	n_PHASE_LOWER:
		lr_ToolRz[n_Robot] := lr_ToolRz[n_Robot] * (1.0 - MIN(1.0, lr_Dt * 5.0));
		IF n_Robot = 1 THEN
			lr_TiltRx := _FC_DemoApproach(lr_TiltRx, 0, lr_TILT_SPEED * lr_Dt);
		END_IF
		(* Delta 2 puts the product down straight (both operands are evaluated). *)
		IF m_MoveToward(vio_Tcp := Tcp[n_Robot], vi_lr_TargetX := Tcp[n_Robot].fX, vi_lr_TargetY := Tcp[n_Robot].fY,
			vi_lr_TargetZ := DEMO_GlobalConst.DEMO_lr_BELT_Z + lr_HeldHeight + lr_GripHeight,
			vi_lr_MaxStep := lr_Step)
		AND (n_Robot <> 1 OR lr_TiltRx = 0)
		THEN
			n_Phase[n_Robot] := n_PHASE_RELEASE;
		END_IF

	n_PHASE_RELEASE:
		(* Every carried product is put down where its finger (Delta 3: the flange) holds it. *)
		FOR n_Slot := 0 TO n_HeldCount[n_Robot] - 1 DO
			IF n_HeldBelt[n_Robot, n_Slot] = 0 THEN
				fb_RefBelt REF= fb_Infeed1;
			ELSE
				fb_RefBelt REF= fb_Infeed2;
			END_IF
			(* Put down on the outfeed: it no longer lies on the infeed. *)
			fb_RefBelt.m_RemoveProduct(udn_Held[n_Robot, n_Slot]);
			n_Finger := SEL(n_Robot = 2, n_Slot + 1, 0);
			Grip := m_GripOffset(vi_n_Robot := n_Robot, vi_n_Finger := n_Finger);
			LatchPose.fX := Tcp[n_Robot].fX + Grip.fX;
			LatchPose.fY := Tcp[n_Robot].fY + Grip.fY;
			LatchPose.fZ := DEMO_GlobalConst.DEMO_lr_BELT_Z;
			(* A product carried at a finger keeps the finger's turn; one at the flange is turned with the base. *)
			LatchPose.fRz := SEL(n_Robot = 2, lr_ToolRz[n_Robot], 0);
			IF fb_Outfeed.m_LatchProduct(vi_udn_Id := DEMO_GlobalVar.DEMO_udn_NextId,
				vi_LatchPose := fb_Outfeed.m_McsToBelt(vi_Pose := LatchPose),
				vi_udn_ProductType := udn_HeldType[n_Robot, n_Slot], vi_lr_LatchBeltPosition := 0,
				vi_b_UseLatchBeltPosition := FALSE, vi_e_State := E_VisuProductState.PLACED,
				vi_udn_ClientId := fb_RefRobot.m_Id())
			THEN
				(* A sample stays marked on the outfeed. *)
				fb_Outfeed.m_SetProductMark(vi_udn_Id := DEMO_GlobalVar.DEMO_udn_NextId, vi_un_Mark := un_HeldMark[n_Robot, n_Slot]);
				DEMO_GlobalVar.DEMO_udn_NextId := DEMO_GlobalVar.DEMO_udn_NextId + 1;
			END_IF
			udn_Held[n_Robot, n_Slot] := 0;
		END_FOR
		n_HeldCount[n_Robot] := 0;
		un_Placed[n_Robot] := un_Placed[n_Robot] + 1;
		n_Phase[n_Robot] := n_PHASE_IDLE;
END_CASE
m_Sequence := TRUE;
END_METHOD

(****************************************************************************************************<br>
© Syntegon Group.<br>
All rights reserved, also regarding any disposal, exploitation, reproduction, editing, distribution,<br>
as well as in the event of applications for industrial property rights.<br>
*****************************************************************************************************<br>
DESCRIPTION:<br>
Follows the current target of Delta n_Robot by its id (register indices shift when entries are removed),<br>
selects its infeed into fb_RefBelt and the finger used for the current pick into n_Finger and Grip. Sets the height<br>
of the product carried or approached and the Delta 3 finger distance closed around it.<br>
****************************************************************************************************)
METHOD PRIVATE m_Target : BOOL
VAR
	lr_TempHalfLength					: LREAL;	// [mm]
	lr_TempHalfWidth					: LREAL;	// [mm]
	lr_TempRadius						: LREAL;	// [mm] corner radius of a rounded box
	lr_TempOuter						: LREAL;	// [mm] radius of the circle around the product's outline
END_VAR
(* Current target *)
b_Found := FALSE;
IF udn_TargetId[n_Robot] <> 0 THEN
	IF n_TargetBelt[n_Robot] = 0 THEN
		fb_RefBelt REF= fb_Infeed1;
	ELSE
		fb_RefBelt REF= fb_Infeed2;
	END_IF
	IF fb_RefBelt.m_FindProduct(udn_TargetId[n_Robot]) >= 0 THEN
		b_Found := fb_RefBelt.m_GetProduct(vi_un_Index := INT_TO_UINT(fb_RefBelt.m_FindProduct(udn_TargetId[n_Robot])),
			vo_Product => Product, vo_Pose => ProductPose);
	END_IF
END_IF

(* Only approaching and descending follow a target; carried products are tracked in udn_Held. *)
IF (n_Phase[n_Robot] = n_PHASE_APPROACH OR n_Phase[n_Robot] = n_PHASE_DESCEND) AND NOT b_Found THEN
	n_Phase[n_Robot] := n_PHASE_IDLE;
	udn_TargetId[n_Robot] := 0;
END_IF
IF b_Found THEN
	ProductPose := fb_RefBelt.m_BeltToMcs(vi_Pose := ProductPose);
	lr_X := ProductPose.fX + lr_LEAD;
	lr_Y := ProductPose.fY;
	lr_TopZ := ProductPose.fZ + lr_TYPE_HEIGHT[LIMIT(1, Product.nProductType, udn_TYPE_COUNT)];
	lr_TargetRz := ProductPose.fRz;
END_IF

(* Size of the product carried, else of the one approached: Delta 1 carries a pair of one type, so its first slot
   stands for both. *)
IF n_HeldCount[n_Robot] > 0 THEN
	udn_Type := LIMIT(1, udn_HeldType[n_Robot, 0], udn_TYPE_COUNT);
ELSIF b_Found THEN
	udn_Type := LIMIT(1, Product.nProductType, udn_TYPE_COUNT);
ELSE
	udn_Type := 1;
END_IF
lr_HeldHeight := lr_TYPE_HEIGHT[udn_Type];
(* Delta 3 closes its fingers on a circle just around the product's outline: around a box's corners, a cylinder's
   larger radius, or a rounded box's corner arcs. *)
lr_TempHalfLength := lr_TYPE_LENGTH[udn_Type] / 2.0;
lr_TempHalfWidth := lr_TYPE_WIDTH[udn_Type] / 2.0;
CASE e_TYPE_SHAPE[udn_Type] OF
	E_VisuProductShape.CYLINDER:
		lr_TempOuter := MAX(lr_TempHalfLength, lr_TempHalfWidth);
	E_VisuProductShape.ROUNDED_BOX:
		lr_TempRadius := MIN(lr_TYPE_CORNER_RADIUS[udn_Type], MIN(lr_TempHalfLength, lr_TempHalfWidth));
		lr_TempOuter := SQRT((lr_TempHalfLength - lr_TempRadius) * (lr_TempHalfLength - lr_TempRadius)
							+ (lr_TempHalfWidth - lr_TempRadius) * (lr_TempHalfWidth - lr_TempRadius)) + lr_TempRadius;
ELSE
	lr_TempOuter := SQRT(lr_TempHalfLength * lr_TempHalfLength + lr_TempHalfWidth * lr_TempHalfWidth);
END_CASE
lr_SpreadClosed := lr_TempOuter + lr_RING_CLEARANCE;

(* Finger used for the current pick: Delta 1 fills its cups one after the other, Delta 3 carries at the flange
   between its fingers. *)
CASE n_Robot OF
	0:
		n_Finger := MIN(n_HeldCount[n_Robot] + 1, 2);
		lr_GripHeight := DEMO_GlobalConst.DEMO_lr_CUP_HEIGHT;
	1:
		n_Finger := 1;
		lr_GripHeight := lr_TILT_HEIGHT;
ELSE
	n_Finger := 0;
	lr_GripHeight := 0;
END_CASE
Grip := m_GripOffset(vi_n_Robot := n_Robot, vi_n_Finger := n_Finger);
m_Target := b_Found;
END_METHOD

(****************************************************************************************************<br>
© Syntegon Group.<br>
All rights reserved, also regarding any disposal, exploitation, reproduction, editing, distribution,<br>
as well as in the event of applications for industrial property rights.<br>
*****************************************************************************************************<br>
DESCRIPTION:<br>
The demo's tracking of Vision 1: latches a raw detection on Infeed 1 at the belt position it was seen at, as<br>
Vision 1's, and marks every tenth product as a sample.<br>
*****************************************************************************************************<br>
OUTPUT VALUES:<br>
TRUE if the product entered the register.<br>
****************************************************************************************************)
METHOD PRIVATE m_Track : BOOL
VAR_INPUT
	vi_Detection						: TVisuDemo_Detection;	// from the product generator
END_VAR
m_Track := fb_Infeed1.m_LatchProduct(vi_udn_Id := DEMO_GlobalVar.DEMO_udn_NextId,
	vi_LatchPose := fb_Infeed1.m_McsToBelt(vi_Pose := vi_Detection.Pose),
	vi_udn_ProductType := vi_Detection.udn_ProductType, vi_lr_LatchBeltPosition := vi_Detection.lr_BeltPosition,
	vi_b_UseLatchBeltPosition := TRUE, vi_e_State := E_VisuProductState.DETECTED, vi_udn_ClientId := fb_Vision1.m_Id());
IF m_Track THEN
	un_Vision1Latches := un_Vision1Latches + 1;
	IF un_Vision1Latches MOD un_SAMPLE_EVERY = 0 THEN
		fb_Infeed1.m_SetProductMark(vi_udn_Id := DEMO_GlobalVar.DEMO_udn_NextId, vi_un_Mark := un_SAMPLE_MARK);
	END_IF
	DEMO_GlobalVar.DEMO_udn_NextId := DEMO_GlobalVar.DEMO_udn_NextId + 1;
END_IF
END_METHOD

END_PROGRAM

// ---- POUs/P_VisuDemoFxx.TcPOU
(****************************************************************************************************<br>
© Syntegon Group.<br>
All rights reserved, also regarding any disposal, exploitation, reproduction, editing, distribution,<br>
as well as in the event of applications for industrial property rights.<br>
*****************************************************************************************************<br>
DESCRIPTION:<br>
DEMO ONLY: Fxx application (Y = 2500). Products arrive irregularly on the Fxx infeed; an XTS loop above the belts<br>
takes them over and puts them onto the Fxx outfeed with an even spacing. Mover 3 and the first far curve module<br>
are in a fault now and then. The Fxx outfeed is a conveyor without a body.<br>
Called by P_VisuDemo.<br>
****************************************************************************************************)
PROGRAM P_VisuDemoFxx
VAR
	fb_FxxInfeed						: _FB_VisuConveyor;
	fb_FxxOutfeed						: _FB_VisuConveyor;
	fb_Fxx								: _FB_VisuXtsLoop;

	(* Conveyors *)
	lr_Dt								: LREAL;	// [s] cycle time
	udn_Seed							: UDINT := 23456;	// [-] pseudo random generator state
	lr_InfeedPosition					: LREAL;	// [mm] belt position of the Fxx infeed
	lr_OutfeedPosition					: LREAL;	// [mm] belt position of the Fxx outfeed
	lr_SinceSpawn						: LREAL;	// [s] since the last product
	lr_SpawnInterval					: LREAL := 0.6;	// [s] irregular: the Fxx evens the gaps out
	BeltPose							: ST_VisuPose;
	LatchPose							: ST_VisuPlanarPose;
	XtsPose								: ST_VisuPose;

	(* XTS loop: unwrapped track position per mover; queued movers wait just before the perimeter (= 0). *)
	b_LoopInitialised					: BOOL;
	lr_LoopS							: ARRAY[0..11] OF LREAL;	// [mm] per mover (n_LOOP_MOVERS)
	n_LoopMode							: ARRAY[0..11] OF INT;
	udn_LoopProduct						: ARRAY[0..11] OF UDINT;	// [-] product id on the Fxx infeed
	MoverFingers						: ARRAY[0..VISU_GlobalConst_Param.VISU_un_MAX_FINGERS - 1] OF ST_VisuFingerState;	// the mover's cup: grips
	un_Module							: UINT;	// [-] track module being set
	e_ModuleKind						: E_VisuModuleKind;
END_VAR
VAR CONSTANT
	lr_FXX_Y							: LREAL := 2500;	// [mm]
	lr_FXX_INFEED_LENGTH				: LREAL := 2000;	// [mm]
	lr_FXX_INFEED_SPEED					: LREAL := 150;	// [mm/s]
	lr_FXX_OUTFEED_X					: LREAL := 2400;	// [mm]
	lr_FXX_OUTFEED_LENGTH				: LREAL := 3000;	// [mm]
	lr_FXX_OUTFEED_SPEED				: LREAL := 300;	// [mm/s]
	lr_LOOP_X							: LREAL := 1000;	// [mm] start of the lower straight above the Fxx infeed
	un_LOOP_STRAIGHT_MODULES			: UINT := 10;	// [-] straight XTS modules per side, joined at each end by two left curve modules
	lr_LOOP_TOOL_OFFSET					: LREAL := 120;	// [mm]
	n_LOOP_MOVERS						: INT := 12;	// [-] size of the lr_LoopS, n_LoopMode and udn_LoopProduct arrays
	lr_LOOP_SLOT						: LREAL := 130;	// [mm] queue spacing
	lr_LOOP_GRIP						: LREAL := 300;	// [mm] track position where the product is gripped
	lr_LOOP_RELEASE						: LREAL := 600;	// [mm] track position where the mover stops following the infeed
	lr_LOOP_PLACE						: LREAL := 2000;	// [mm] track position of the hand-over to the Fxx outfeed
	lr_LOOP_DELIVER_SPEED				: LREAL := 700;	// [mm/s]
	lr_LOOP_RETURN_SPEED				: LREAL := 900;	// [mm/s]
	lr_FAULT_START						: LREAL := 10;	// [s] start of the mover 3 fault in the fault period
	lr_MODULE_FAULT_START				: LREAL := 15;	// [s] start of the fault of the first far curve module
	n_LOOP_QUEUE						: INT := 0;
	n_LOOP_TRACK						: INT := 1;
	n_LOOP_DELIVER						: INT := 2;
	n_LOOP_RETURN						: INT := 3;
END_VAR

lr_Dt := DEMO_GlobalVar.DEMO_lr_Dt;


(****************************************************************************************************)
(* REGISTRATION (idempotent, every cycle)                                                           *)
(****************************************************************************************************)
fb_FxxInfeed.m_Register(vio_Manifest := GVL_Visu.stManifest, vi_udn_Id := 4, vi_str_Name := 'Fxx infeed');
fb_FxxOutfeed.m_Register(vio_Manifest := GVL_Visu.stManifest, vi_udn_Id := 5, vi_str_Name := 'Fxx outfeed');
fb_Fxx.m_Register(vio_Manifest := GVL_Visu.stManifest, vi_udn_Id := 20, vi_str_Name := 'Fxx');


(****************************************************************************************************)
(* CONVEYORS (configuration idempotent, every cycle)                                                *)
(****************************************************************************************************)
BeltPose.fX := 0;
BeltPose.fY := lr_FXX_Y;
BeltPose.fZ := DEMO_GlobalConst.DEMO_lr_BELT_Z;
fb_FxxInfeed.m_SetPose(vi_Pose := BeltPose);
fb_FxxInfeed.m_Configure(vi_lr_Length := lr_FXX_INFEED_LENGTH,
	vi_lr_Width := DEMO_GlobalConst.DEMO_lr_BELT_WIDTH);
BeltPose.fX := lr_FXX_OUTFEED_X;
(* The outfeed's coordinate system lies on its right edge (seen in the conveying direction). *)
fb_FxxOutfeed.m_SetOriginShift(vi_lr_X := 0, vi_lr_Y := -DEMO_GlobalConst.DEMO_lr_BELT_WIDTH / 2, vi_lr_Z := 0);
fb_FxxOutfeed.m_SetPose(vi_Pose := BeltPose);
fb_FxxOutfeed.m_Configure(vi_lr_Length := lr_FXX_OUTFEED_LENGTH,
	vi_lr_Width := DEMO_GlobalConst.DEMO_lr_BELT_WIDTH);
(* A conveyor without a body: only its products, zones and axis (from the shifted origin) are drawn. *)
fb_FxxOutfeed.m_SetBodyVisible(vi_b_Visible := FALSE);
fb_FxxInfeed.m_SetProductType(vi_udn_Id := 1, vi_lr_Length := DEMO_GlobalConst.DEMO_lr_PRODUCT_LENGTH,
	vi_lr_Width := DEMO_GlobalConst.DEMO_lr_PRODUCT_WIDTH, vi_lr_Height := DEMO_GlobalConst.DEMO_lr_PRODUCT_HEIGHT,
	vi_e_Shape := E_VisuProductShape.BOX, vi_lr_CornerRadius := 0);
fb_FxxOutfeed.m_SetProductType(vi_udn_Id := 1, vi_lr_Length := DEMO_GlobalConst.DEMO_lr_PRODUCT_LENGTH,
	vi_lr_Width := DEMO_GlobalConst.DEMO_lr_PRODUCT_WIDTH, vi_lr_Height := DEMO_GlobalConst.DEMO_lr_PRODUCT_HEIGHT,
	vi_e_Shape := E_VisuProductShape.BOX, vi_lr_CornerRadius := 0);

(* Belt travel *)
lr_InfeedPosition := lr_InfeedPosition + lr_FXX_INFEED_SPEED * lr_Dt;
lr_OutfeedPosition := lr_OutfeedPosition + lr_FXX_OUTFEED_SPEED * lr_Dt;
fb_FxxInfeed.m_SetBeltPosition(lr_InfeedPosition);
fb_FxxOutfeed.m_SetBeltPosition(lr_OutfeedPosition);


(****************************************************************************************************)
(* PRODUCT INFEED: irregular gaps                                                                   *)
(****************************************************************************************************)
lr_SinceSpawn := lr_SinceSpawn + lr_Dt;
IF lr_SinceSpawn >= lr_SpawnInterval THEN
	lr_SinceSpawn := 0;
	udn_Seed := udn_Seed * 1103515245 + 12345;
	lr_SpawnInterval := 0.4 + UDINT_TO_LREAL(udn_Seed MOD 1000) / 1000.0 * 1.2;
	LatchPose.fX := 100;
	LatchPose.fY := lr_FXX_Y;
	LatchPose.fZ := DEMO_GlobalConst.DEMO_lr_BELT_Z;
	LatchPose.fRz := 0;
	IF fb_FxxInfeed.m_LatchProduct(vi_udn_Id := DEMO_GlobalVar.DEMO_udn_NextId,
		vi_LatchPose := fb_FxxInfeed.m_McsToBelt(vi_Pose := LatchPose),
		vi_udn_ProductType := 1, vi_lr_LatchBeltPosition := 0, vi_b_UseLatchBeltPosition := FALSE,
		vi_e_State := E_VisuProductState.DETECTED, vi_udn_ClientId := 0)
	THEN
		DEMO_GlobalVar.DEMO_udn_NextId := DEMO_GlobalVar.DEMO_udn_NextId + 1;
	END_IF
END_IF


(****************************************************************************************************)
(* XTS LOOP                                                                                         *)
(****************************************************************************************************)
XtsPose.fX := lr_LOOP_X;
XtsPose.fY := lr_FXX_Y;
XtsPose.fZ := DEMO_GlobalConst.DEMO_lr_BELT_Z + DEMO_GlobalConst.DEMO_lr_PRODUCT_HEIGHT + lr_LOOP_TOOL_OFFSET;
XtsPose.fRz := 0;
(* The flange sits one cup height closer to the track, so the cup's grip point is at the products' tops. *)
fb_Fxx.m_SetPose(vi_Pose := XtsPose);
fb_Fxx.m_Configure(vi_lr_ToolOffset := lr_LOOP_TOOL_OFFSET - DEMO_GlobalConst.DEMO_lr_CUP_HEIGHT,
	vi_lr_MoverLength := 100, vi_lr_MoverWidth := 60);
(* Track: per side the straight modules, then two left curve modules turning up and back. *)
FOR un_Module := 1 TO 2 * (un_LOOP_STRAIGHT_MODULES + 2) DO
	IF (un_Module - 1) MOD (un_LOOP_STRAIGHT_MODULES + 2) < un_LOOP_STRAIGHT_MODULES THEN
		e_ModuleKind := E_VisuModuleKind.STRAIGHT;
	ELSE
		e_ModuleKind := E_VisuModuleKind.CURVE_LEFT;
	END_IF
	fb_Fxx.m_SetModule(vi_un_Module := un_Module, vi_e_Kind := e_ModuleKind,
		vi_lr_Length := VISU_GlobalConst.VISU_lr_XTS_MODULE_LENGTH);
END_FOR
fb_Fxx.m_SetModuleFault(vi_un_Module := un_LOOP_STRAIGHT_MODULES + 1,
	vi_b_Fault := DEMO_GlobalVar.DEMO_lr_FaultPhase >= lr_MODULE_FAULT_START
					AND DEMO_GlobalVar.DEMO_lr_FaultPhase < lr_MODULE_FAULT_START + DEMO_GlobalConst.DEMO_lr_FAULT_DURATION,
	vi_str_FaultMessage := 'Overtemperature');
fb_Fxx.m_SetFinger(vi_un_Finger := 1, vi_lr_Diameter := DEMO_GlobalConst.DEMO_lr_CUP_DIAMETER,
	vi_lr_Height := DEMO_GlobalConst.DEMO_lr_CUP_HEIGHT);
(* The cup hangs at the flange centre; the movers report no finger poses, the visualisation places the cup by its
   offset on every mover's flange (ADR 0018). *)
fb_Fxx.m_SetFingerOffset(vi_un_Finger := 1, vi_lr_X := 0, vi_lr_Y := 0, vi_lr_Z := 0, vi_lr_Rz := 0);
fb_Fxx.m_SetFingersOnFlange(vi_b_OnFlange := TRUE);
fb_Fxx.m_SetZone(vi_un_Zone := 1, vi_udn_ConveyorId := fb_FxxInfeed.m_Id(), vi_lr_Start := lr_LOOP_X,
	vi_lr_End := lr_LOOP_X + lr_LOOP_RELEASE, vi_lr_AllocationOffset := 0, vi_lr_CcsOffset := lr_LOOP_X,
	vi_lr_StartY := 0, vi_lr_EndY := 0);
fb_Fxx.m_SetZone(vi_un_Zone := 2, vi_udn_ConveyorId := fb_FxxOutfeed.m_Id(),
	vi_lr_Start := lr_LOOP_X + lr_LOOP_PLACE - lr_FXX_OUTFEED_X - 300,
	vi_lr_End := lr_LOOP_X + lr_LOOP_PLACE - lr_FXX_OUTFEED_X + 100,
	vi_lr_AllocationOffset := 0, vi_lr_CcsOffset := lr_LOOP_X + lr_LOOP_PLACE - lr_FXX_OUTFEED_X,
	vi_lr_StartY := 0, vi_lr_EndY := 0);
m_Step();


(****************************************************************************************************)
(* HOUSEKEEPING                                                                                     *)
(****************************************************************************************************)
fb_FxxInfeed.m_RemoveProductsBeyond(lr_FXX_INFEED_LENGTH + DEMO_GlobalConst.DEMO_lr_REMOVE_BEYOND_END);
fb_FxxOutfeed.m_RemoveProductsBeyond(lr_FXX_OUTFEED_LENGTH + DEMO_GlobalConst.DEMO_lr_REMOVE_BEYOND_END);

(****************************************************************************************************<br>
© Syntegon Group.<br>
All rights reserved, also regarding any disposal, exploitation, reproduction, editing, distribution,<br>
as well as in the event of applications for industrial property rights.<br>
*****************************************************************************************************<br>
DESCRIPTION:<br>
XTS loop: the queue head takes over the next product arriving on the Fxx infeed under the start of the lower<br>
straight, follows it, grips it, carries it faster to the Fxx outfeed and releases it there; the mover then<br>
runs round to the queue.<br>
****************************************************************************************************)
METHOD PRIVATE m_Step : BOOL
VAR
	lr_TempPerimeter					: LREAL;	// [mm]
	lr_TempS							: LREAL;	// [mm]
	lr_TempX							: LREAL;	// [mm]
	lr_TempRz							: LREAL;	// [deg]
	n_TempI								: INT;
	n_TempJ								: INT;
	n_TempRank							: INT;
	n_TempHead							: INT;
	b_TempHeadReady						: BOOL;
	lr_TempMinTrack						: LREAL;	// [mm]
	n_TempIdx							: INT;
	un_TempIndex						: UINT;
	TempProduct							: ST_VisuProduct;
	TempPose							: ST_VisuPlanarPose;
	TempLatch							: ST_VisuPlanarPose;
END_VAR
(****************************************************************************************************)
(* QUEUE AND TAKE-OVER                                                                              *)
(****************************************************************************************************)
lr_TempPerimeter := fb_Fxx.m_TrackLength();
IF NOT b_LoopInitialised THEN
	FOR n_TempI := 0 TO n_LOOP_MOVERS - 1 DO
		lr_LoopS[n_TempI] := lr_TempPerimeter - INT_TO_LREAL(n_TempI) * lr_LOOP_SLOT;
		n_LoopMode[n_TempI] := n_LOOP_QUEUE;
	END_FOR
	b_LoopInitialised := TRUE;
END_IF

(* Queued movers close up towards their slots before the start of the lower straight. *)
n_TempHead := -1;
FOR n_TempI := 0 TO n_LOOP_MOVERS - 1 DO
	IF n_LoopMode[n_TempI] = n_LOOP_QUEUE THEN
		n_TempRank := 0;
		FOR n_TempJ := 0 TO n_LOOP_MOVERS - 1 DO
			IF n_LoopMode[n_TempJ] = n_LOOP_QUEUE
			AND (lr_LoopS[n_TempJ] > lr_LoopS[n_TempI] OR (lr_LoopS[n_TempJ] = lr_LoopS[n_TempI] AND n_TempJ < n_TempI))
			THEN
				n_TempRank := n_TempRank + 1;
			END_IF
		END_FOR
		lr_LoopS[n_TempI] := MIN(lr_LoopS[n_TempI] + lr_LOOP_RETURN_SPEED * lr_Dt,
								lr_TempPerimeter - INT_TO_LREAL(n_TempRank) * lr_LOOP_SLOT);
		IF n_TempRank = 0 THEN
			n_TempHead := n_TempI;
		END_IF
	END_IF
END_FOR

(* The queue head takes over the next product arriving under the start of the lower straight.
   ST evaluates both operands of AND, so the index check must be a separate IF (head = -1: queue empty). *)
b_TempHeadReady := FALSE;
IF n_TempHead >= 0 THEN
	b_TempHeadReady := lr_LoopS[n_TempHead] >= lr_TempPerimeter - 1;
END_IF
(* Movers cannot overlap: the next product must be at least one slot behind the last mover following one. *)
lr_TempMinTrack := 1.0E9;
FOR n_TempI := 0 TO n_LOOP_MOVERS - 1 DO
	IF n_LoopMode[n_TempI] = n_LOOP_TRACK THEN
		lr_TempMinTrack := MIN(lr_TempMinTrack, lr_LoopS[n_TempI]);
	END_IF
END_FOR
IF b_TempHeadReady THEN
	un_TempIndex := 0;
	WHILE n_LoopMode[n_TempHead] = n_LOOP_QUEUE AND un_TempIndex < fb_FxxInfeed.m_ProductCount() DO
		fb_FxxInfeed.m_GetProduct(vi_un_Index := un_TempIndex, vo_Product => TempProduct, vo_Pose => TempPose);
		TempPose := fb_FxxInfeed.m_BeltToMcs(vi_Pose := TempPose);
		lr_TempX := TempPose.fX - lr_LOOP_X;
		IF TempProduct.eState = E_VisuProductState.DETECTED AND lr_TempX >= 0 AND lr_TempX < lr_LOOP_GRIP
		AND lr_TempMinTrack - lr_TempX >= lr_LOOP_SLOT
		THEN
			fb_FxxInfeed.m_SetProductState(vi_udn_Id := TempProduct.nId, vi_e_State := E_VisuProductState.ASSIGNED,
				vi_udn_ClientId := fb_Fxx.m_Id(), vi_udn_MoverId := INT_TO_UDINT(n_TempHead + 1), vi_udn_FingerId := 0);
			udn_LoopProduct[n_TempHead] := TempProduct.nId;
			n_LoopMode[n_TempHead] := n_LOOP_TRACK;
		END_IF
		un_TempIndex := un_TempIndex + 1;
	END_WHILE
END_IF


(****************************************************************************************************)
(* MOVERS                                                                                           *)
(****************************************************************************************************)
fb_Fxx.m_SetMoverCount(INT_TO_UINT(n_LOOP_MOVERS));
FOR n_TempI := 0 TO n_LOOP_MOVERS - 1 DO
	CASE n_LoopMode[n_TempI] OF
		n_LOOP_TRACK:
			n_TempIdx := fb_FxxInfeed.m_FindProduct(udn_LoopProduct[n_TempI]);
			IF n_TempIdx < 0 THEN
				udn_LoopProduct[n_TempI] := 0;
				n_LoopMode[n_TempI] := n_LOOP_RETURN;
			ELSE
				fb_FxxInfeed.m_GetProduct(vi_un_Index := INT_TO_UINT(n_TempIdx), vo_Product => TempProduct, vo_Pose => TempPose);
				TempPose := fb_FxxInfeed.m_BeltToMcs(vi_Pose := TempPose);
				lr_LoopS[n_TempI] := TempPose.fX - lr_LOOP_X;
				IF lr_LoopS[n_TempI] >= lr_LOOP_GRIP AND TempProduct.eState = E_VisuProductState.ASSIGNED THEN
					fb_FxxInfeed.m_SetProductState(vi_udn_Id := TempProduct.nId, vi_e_State := E_VisuProductState.PICKED,
						vi_udn_ClientId := fb_Fxx.m_Id(), vi_udn_MoverId := INT_TO_UDINT(n_TempI + 1), vi_udn_FingerId := 1);
				END_IF
				IF lr_LoopS[n_TempI] >= lr_LOOP_RELEASE THEN
					n_LoopMode[n_TempI] := n_LOOP_DELIVER;
				END_IF
			END_IF

		n_LOOP_DELIVER:
			lr_LoopS[n_TempI] := MIN(lr_LoopS[n_TempI] + lr_LOOP_DELIVER_SPEED * lr_Dt, lr_LOOP_PLACE);
			IF lr_LoopS[n_TempI] >= lr_LOOP_PLACE THEN
				lr_TempRz := 0;
				n_TempIdx := fb_FxxInfeed.m_FindProduct(udn_LoopProduct[n_TempI]);
				IF n_TempIdx >= 0 THEN
					fb_FxxInfeed.m_GetProduct(vi_un_Index := INT_TO_UINT(n_TempIdx), vo_Product => TempProduct, vo_Pose => TempPose);
					lr_TempRz := TempProduct.stLatchPose.fRz;
					(* Put down on the outfeed: it no longer lies on the infeed. *)
					fb_FxxInfeed.m_RemoveProduct(TempProduct.nId);
				END_IF
				TempLatch.fX := lr_LOOP_X + lr_LoopS[n_TempI];
				TempLatch.fY := lr_FXX_Y;
				TempLatch.fZ := DEMO_GlobalConst.DEMO_lr_BELT_Z;
				TempLatch.fRz := lr_TempRz;
				IF fb_FxxOutfeed.m_LatchProduct(vi_udn_Id := DEMO_GlobalVar.DEMO_udn_NextId,
					vi_LatchPose := fb_FxxOutfeed.m_McsToBelt(vi_Pose := TempLatch),
					vi_udn_ProductType := 1, vi_lr_LatchBeltPosition := 0, vi_b_UseLatchBeltPosition := FALSE,
					vi_e_State := E_VisuProductState.PLACED, vi_udn_ClientId := fb_Fxx.m_Id())
				THEN
					DEMO_GlobalVar.DEMO_udn_NextId := DEMO_GlobalVar.DEMO_udn_NextId + 1;
				END_IF
				udn_LoopProduct[n_TempI] := 0;
				n_LoopMode[n_TempI] := n_LOOP_RETURN;
			END_IF

		n_LOOP_RETURN:
			lr_LoopS[n_TempI] := lr_LoopS[n_TempI] + lr_LOOP_RETURN_SPEED * lr_Dt;
			IF lr_LoopS[n_TempI] >= lr_TempPerimeter - INT_TO_LREAL(n_LOOP_MOVERS) * lr_LOOP_SLOT THEN
				n_LoopMode[n_TempI] := n_LOOP_QUEUE;
			END_IF
	END_CASE

	(* Report the mover with its cup: whether it grips; its pose follows from its offset on the flange. *)
	lr_TempS := lr_LoopS[n_TempI];
	IF lr_TempS >= lr_TempPerimeter THEN
		lr_TempS := lr_TempS - lr_TempPerimeter;
	END_IF
	MoverFingers[0].bActive := n_LoopMode[n_TempI] = n_LOOP_DELIVER
							OR (n_LoopMode[n_TempI] = n_LOOP_TRACK AND lr_LoopS[n_TempI] >= lr_LOOP_GRIP);

	(* Demo fault: mover 3 now and then. *)
	fb_Fxx.m_SetMover(vi_un_Index := INT_TO_UINT(n_TempI), vi_udn_Id := INT_TO_UDINT(n_TempI + 1), vi_lr_Position := lr_TempS,
		vi_FingerStates := MoverFingers,
		vi_b_Fault := n_TempI = 2 AND DEMO_GlobalVar.DEMO_lr_FaultPhase >= lr_FAULT_START
					AND DEMO_GlobalVar.DEMO_lr_FaultPhase < lr_FAULT_START + DEMO_GlobalConst.DEMO_lr_FAULT_DURATION,
		vi_str_FaultMessage := 'Following error');
END_FOR
m_Step := TRUE;
END_METHOD

END_PROGRAM

// ---- POUs/P_VisuDemoIdh.TcPOU
(****************************************************************************************************<br>
© Syntegon Group.<br>
All rights reserved, also regarding any disposal, exploitation, reproduction, editing, distribution,<br>
as well as in the event of applications for industrial property rights.<br>
*****************************************************************************************************<br>
DESCRIPTION:<br>
DEMO ONLY: IDH application (Y = 4100..4850). An XTS gantry with four movers picks products from the IDH infeed<br>
in batches and places them onto the tray belt. Mover 2 is in a fault now and then. Called by P_VisuDemo.<br>
****************************************************************************************************)
PROGRAM P_VisuDemoIdh
VAR
	fb_IdhInfeed						: _FB_VisuConveyor;
	fb_IdhTray							: _FB_VisuConveyor;
	fb_Idh								: _FB_VisuXtsGantry;
	(* Syn_Config (ADR 0017): the IDH runs with the parameter set the configurator writes (pose, track, zones,
	   gripper, limit areas), else with its program values; taken over at once in the demo. The simulated motion keeps to the
	   program's track. *)
	fb_IdhParam							: SynConfig._FB_ConfigXtsGantry;
	IdhDefault							: SynConfig.ST_ConfigXtsGantryParam;	// program values of the IDH

	(* Conveyors *)
	lr_Dt								: LREAL;	// [s] cycle time
	udn_Seed							: UDINT := 34567;	// [-] pseudo random generator state
	lr_InfeedPosition					: LREAL;	// [mm] belt position of the IDH infeed
	lr_TrayPosition						: LREAL;	// [mm] belt position of the tray belt
	lr_SinceSpawn						: LREAL;	// [s] since the last product
	lr_SpawnInterval					: LREAL := 0.8;	// [s]
	BeltPose							: ST_VisuPose;
	LatchPose							: ST_VisuPlanarPose;

	(* XTS gantry *)
	n_GantryPhase						: INT;
	lr_GantryZ							: LREAL;	// [mm]
	lr_GantryWait						: ARRAY[0..3] OF LREAL := [100, 300, 500, 700];	// [mm]
	lr_GantryPos						: ARRAY[0..3] OF LREAL := [100, 300, 500, 700];	// [mm]
	lr_GantryX							: ARRAY[0..3] OF LREAL := [200, 200, 200, 200];	// [mm]
	lr_GantryC							: ARRAY[0..3] OF LREAL;	// [deg]
	b_GantryGrip						: ARRAY[0..3] OF BOOL;
	udn_GantryProduct					: ARRAY[0..3] OF UDINT;	// [-] product id on the IDH infeed
	MoverFingers						: ARRAY[0..VISU_GlobalConst_Param.VISU_un_MAX_FINGERS - 1] OF ST_VisuFingerState;	// the mover's cup
	un_Module							: UINT;	// [-] track module being set
END_VAR
VAR PERSISTENT
	IdhSet								: SynConfig.ST_ConfigXtsGantrySet;	// active parameter set of the IDH, kept over a restart
END_VAR
VAR CONSTANT
	(* Gantry turned by -90 deg: track along MCS +X, X axes towards MCS -Y (IDH infeed under X = 200, tray belt
	   under X = 600). *)
	lr_IDH_INFEED_Y						: LREAL := 4500;	// [mm]
	lr_IDH_INFEED_LENGTH				: LREAL := 4000;	// [mm]
	lr_IDH_INFEED_SPEED					: LREAL := 200;	// [mm/s]
	lr_TRAY_X							: LREAL := 1300;	// [mm]
	lr_TRAY_Y							: LREAL := 4100;	// [mm]
	lr_TRAY_LENGTH						: LREAL := 2000;	// [mm]
	lr_TRAY_SPEED						: LREAL := 80;	// [mm/s]
	lr_GANTRY_X							: LREAL := 1500;	// [mm]
	lr_GANTRY_Y							: LREAL := 4850;	// [mm]
	lr_GANTRY_Z							: LREAL := 1340;	// [mm]
	un_GANTRY_MODULES					: UINT := 6;	// [-]
	lr_GANTRY_MODULE_LENGTH				: LREAL := 250;	// [mm]
	lr_GANTRY_TOOL_X					: LREAL := 150;	// [mm]
	lr_GANTRY_TOOL_Z					: LREAL := -400;	// [mm]
	lr_GANTRY_MOVER_LENGTH				: LREAL := 155;	// [mm]
	lr_GANTRY_GAP						: LREAL := 180;	// [mm] minimum distance between movers
	lr_GANTRY_X_BELT					: LREAL := 200;	// [mm]
	lr_GANTRY_X_TRAY					: LREAL := 600;	// [mm]
	lr_GANTRY_Z_DOWN					: LREAL := -100;	// [mm]
	lr_GANTRY_Z_SPEED					: LREAL := 500;	// [mm/s]
	lr_GANTRY_X_SPEED					: LREAL := 1000;	// [mm/s]
	lr_GANTRY_TRACK_SPEED				: LREAL := 1500;	// [mm/s]
	lr_FAULT_START						: LREAL := 12;	// [s] start of the mover 2 fault in the fault period
	n_GANTRY_COLLECT					: INT := 0;
	n_GANTRY_PICK_DOWN					: INT := 1;
	n_GANTRY_PICK_UP					: INT := 2;
	n_GANTRY_TO_TRAY					: INT := 3;
	n_GANTRY_PLACE_DOWN					: INT := 4;
	n_GANTRY_PLACE_UP					: INT := 5;
	n_GANTRY_RETURN						: INT := 6;
END_VAR

lr_Dt := DEMO_GlobalVar.DEMO_lr_Dt;


(****************************************************************************************************)
(* REGISTRATION (idempotent, every cycle)                                                           *)
(****************************************************************************************************)
fb_IdhInfeed.m_Register(vio_Manifest := GVL_Visu.stManifest, vi_udn_Id := 6, vi_str_Name := 'IDH infeed');
fb_IdhTray.m_Register(vio_Manifest := GVL_Visu.stManifest, vi_udn_Id := 7, vi_str_Name := 'Tray belt');
fb_Idh.m_Register(vio_Manifest := GVL_Visu.stManifest, vi_udn_Id := 30, vi_str_Name := 'IDH');


(****************************************************************************************************)
(* CONVEYORS (configuration idempotent, every cycle)                                                *)
(****************************************************************************************************)
BeltPose.fX := 0;
BeltPose.fY := lr_IDH_INFEED_Y;
BeltPose.fZ := DEMO_GlobalConst.DEMO_lr_BELT_Z;
fb_IdhInfeed.m_SetPose(vi_Pose := BeltPose);
fb_IdhInfeed.m_Configure(vi_lr_Length := lr_IDH_INFEED_LENGTH,
	vi_lr_Width := DEMO_GlobalConst.DEMO_lr_BELT_WIDTH);
BeltPose.fX := lr_TRAY_X;
BeltPose.fY := lr_TRAY_Y;
fb_IdhTray.m_SetPose(vi_Pose := BeltPose);
fb_IdhTray.m_Configure(vi_lr_Length := lr_TRAY_LENGTH, vi_lr_Width := DEMO_GlobalConst.DEMO_lr_BELT_WIDTH);
fb_IdhInfeed.m_SetProductType(vi_udn_Id := 1, vi_lr_Length := DEMO_GlobalConst.DEMO_lr_PRODUCT_LENGTH,
	vi_lr_Width := DEMO_GlobalConst.DEMO_lr_PRODUCT_WIDTH, vi_lr_Height := DEMO_GlobalConst.DEMO_lr_PRODUCT_HEIGHT,
	vi_e_Shape := E_VisuProductShape.BOX, vi_lr_CornerRadius := 0);
fb_IdhTray.m_SetProductType(vi_udn_Id := 1, vi_lr_Length := DEMO_GlobalConst.DEMO_lr_PRODUCT_LENGTH,
	vi_lr_Width := DEMO_GlobalConst.DEMO_lr_PRODUCT_WIDTH, vi_lr_Height := DEMO_GlobalConst.DEMO_lr_PRODUCT_HEIGHT,
	vi_e_Shape := E_VisuProductShape.BOX, vi_lr_CornerRadius := 0);

(* Belt travel *)
lr_InfeedPosition := lr_InfeedPosition + lr_IDH_INFEED_SPEED * lr_Dt;
lr_TrayPosition := lr_TrayPosition + lr_TRAY_SPEED * lr_Dt;
fb_IdhInfeed.m_SetBeltPosition(lr_InfeedPosition);
fb_IdhTray.m_SetBeltPosition(lr_TrayPosition);


(****************************************************************************************************)
(* PRODUCT INFEED: slightly irregular gaps, products turned                                         *)
(****************************************************************************************************)
lr_SinceSpawn := lr_SinceSpawn + lr_Dt;
IF lr_SinceSpawn >= lr_SpawnInterval THEN
	lr_SinceSpawn := 0;
	udn_Seed := udn_Seed * 1103515245 + 12345;
	lr_SpawnInterval := 0.6 + UDINT_TO_LREAL(udn_Seed MOD 1000) / 1000.0 * 0.6;
	LatchPose.fX := 100;
	LatchPose.fY := lr_IDH_INFEED_Y;
	LatchPose.fZ := DEMO_GlobalConst.DEMO_lr_BELT_Z;
	LatchPose.fRz := (UDINT_TO_LREAL((udn_Seed / 1000) MOD 1000) / 1000.0 - 0.5) * 60.0;
	IF fb_IdhInfeed.m_LatchProduct(vi_udn_Id := DEMO_GlobalVar.DEMO_udn_NextId,
		vi_LatchPose := fb_IdhInfeed.m_McsToBelt(vi_Pose := LatchPose),
		vi_udn_ProductType := 1, vi_lr_LatchBeltPosition := 0, vi_b_UseLatchBeltPosition := FALSE,
		vi_e_State := E_VisuProductState.DETECTED, vi_udn_ClientId := 0)
	THEN
		DEMO_GlobalVar.DEMO_udn_NextId := DEMO_GlobalVar.DEMO_udn_NextId + 1;
	END_IF
END_IF


(****************************************************************************************************)
(* XTS GANTRY                                                                                       *)
(****************************************************************************************************)
(* The IDH's program values; its parameter set (Syn_Config) replaces them once the configurator wrote one. Strokes,
   tool offsets and mover size are hardware and stay the program's. *)
IdhDefault.stPose.fX := lr_GANTRY_X;
IdhDefault.stPose.fY := lr_GANTRY_Y;
IdhDefault.stPose.fZ := lr_GANTRY_Z;
IdhDefault.stPose.fRz := -90;
IdhDefault.nModuleCount := un_GANTRY_MODULES;
FOR un_Module := 1 TO un_GANTRY_MODULES DO
	IdhDefault.aModules[un_Module - 1].eKind := E_VisuModuleKind.STRAIGHT;
	IdhDefault.aModules[un_Module - 1].fLength := lr_GANTRY_MODULE_LENGTH;
END_FOR
(* Limit area in the gantry frame (flange coordinates): around the flanges' travel, from over the infeed to over
   the tray belt, along the whole track. *)
IdhDefault.stLimitArea.fXMin := 250;
IdhDefault.stLimitArea.fXMax := 850;
IdhDefault.stLimitArea.fYMin := -50;
IdhDefault.stLimitArea.fYMax := 1550;
IdhDefault.stLimitArea.fZMin := -600;
IdhDefault.stLimitArea.fZMax := -300;
IdhDefault.stLimitArea.bActive := TRUE;
(* Around every mover's flange, cup and product; narrower along the track than the movers' least distance. *)
IdhDefault.stTcpLimitArea.fXMin := -60;
IdhDefault.stTcpLimitArea.fXMax := 60;
IdhDefault.stTcpLimitArea.fYMin := -85;
IdhDefault.stTcpLimitArea.fYMax := 85;
IdhDefault.stTcpLimitArea.fZMin := -100;
IdhDefault.stTcpLimitArea.fZMax := 20;
IdhDefault.stTcpLimitArea.bActive := TRUE;
IdhDefault.nZoneCount := 2;
IdhDefault.aZones[0].nConveyorId := fb_IdhInfeed.m_Id();
IdhDefault.aZones[0].fStart := lr_GANTRY_X;
IdhDefault.aZones[0].fEnd := lr_GANTRY_X + UINT_TO_LREAL(un_GANTRY_MODULES) * lr_GANTRY_MODULE_LENGTH;
IdhDefault.aZones[0].fCcsOffset := lr_GANTRY_X;
IdhDefault.aZones[1].nConveyorId := fb_IdhTray.m_Id();
IdhDefault.aZones[1].fStart := lr_GANTRY_X - lr_TRAY_X;
IdhDefault.aZones[1].fEnd := lr_GANTRY_X - lr_TRAY_X + UINT_TO_LREAL(un_GANTRY_MODULES) * lr_GANTRY_MODULE_LENGTH;
IdhDefault.aZones[1].fCcsOffset := lr_GANTRY_X - lr_TRAY_X;
(* Every mover's suction cup, at the flange centre (ADR 0018); the movers report its live pose, turned by C. It
   comes with the parameter set: the application no longer calls m_SetFinger itself. *)
IdhDefault.nFingerCount := 1;
IdhDefault.aFingers[0].fDiameter := DEMO_GlobalConst.DEMO_lr_CUP_DIAMETER;
IdhDefault.aFingers[0].fHeight := DEMO_GlobalConst.DEMO_lr_CUP_HEIGHT;
fb_IdhParam.m_Register(vio_Manifest := GVL_Config.stManifest, vi_udn_Id := fb_Idh.m_Id());
fb_IdhParam.m_Cycle(vio_Default := IdhDefault, vio_Set := IdhSet, vi_b_ApplyAllowed := TRUE);
fb_Idh.m_Configure(vi_lr_XMin := 0, vi_lr_XMax := 700, vi_lr_ZMin := lr_GANTRY_Z_DOWN, vi_lr_ZMax := 0,
	vi_lr_ToolOffsetX := lr_GANTRY_TOOL_X, vi_lr_ToolOffsetZ := lr_GANTRY_TOOL_Z + DEMO_GlobalConst.DEMO_lr_CUP_HEIGHT,
	vi_lr_MoverLength := lr_GANTRY_MOVER_LENGTH, vi_lr_MoverWidth := 80);
fb_IdhParam.m_PassOn(vio_Visu := fb_Idh);
m_Step();


(****************************************************************************************************)
(* HOUSEKEEPING                                                                                     *)
(****************************************************************************************************)
fb_IdhInfeed.m_RemoveProductsBeyond(lr_IDH_INFEED_LENGTH + DEMO_GlobalConst.DEMO_lr_REMOVE_BEYOND_END);
fb_IdhTray.m_RemoveProductsBeyond(lr_TRAY_LENGTH + DEMO_GlobalConst.DEMO_lr_REMOVE_BEYOND_END);

(****************************************************************************************************<br>
© Syntegon Group.<br>
All rights reserved, also regarding any disposal, exploitation, reproduction, editing, distribution,<br>
as well as in the event of applications for industrial property rights.<br>
*****************************************************************************************************<br>
DESCRIPTION:<br>
Moves the gantry movers along the track: a mover with a product waits at its waiting position until the<br>
product passes underneath and then follows it; a mover without one returns to its waiting position.<br>
Downstream first, so each mover keeps its distance to the one ahead.<br>
****************************************************************************************************)
METHOD PRIVATE m_Follow : BOOL
VAR
	n_TempI								: INT;
	lr_TempGoal							: LREAL;	// [mm]
	lr_TempLimit						: LREAL;	// [mm]
	lr_TempPos							: LREAL;	// [mm]
	lr_TempRz							: LREAL;	// [deg]
END_VAR
FOR n_TempI := 3 TO 0 BY -1 DO
	IF n_TempI = 3 THEN
		lr_TempLimit := UINT_TO_LREAL(un_GANTRY_MODULES) * lr_GANTRY_MODULE_LENGTH - lr_GANTRY_MOVER_LENGTH / 2;
	ELSE
		lr_TempLimit := lr_GantryPos[n_TempI + 1] - lr_GANTRY_GAP;
	END_IF
	lr_TempGoal := lr_GantryWait[n_TempI];
	IF udn_GantryProduct[n_TempI] <> 0 THEN
		IF m_TrackPos(vi_udn_Id := udn_GantryProduct[n_TempI], vo_lr_TrackPos => lr_TempPos, vo_lr_Rz => lr_TempRz) THEN
			lr_TempGoal := MAX(lr_TempPos, lr_GantryWait[n_TempI]);
			(* The cup turns by -90 + C in the MCS (gantry turned by -90 deg), so C = Rz + 90 meets the product. *)
			lr_GantryC[n_TempI] := _FC_DemoApproach(lr_GantryC[n_TempI], lr_TempRz + 90.0, 180.0 * lr_Dt);
		END_IF
	END_IF
	lr_GantryPos[n_TempI] := MIN(_FC_DemoApproach(lr_GantryPos[n_TempI], lr_TempGoal, lr_GANTRY_TRACK_SPEED * lr_Dt),
								lr_TempLimit);
END_FOR
m_Follow := TRUE;
END_METHOD

(****************************************************************************************************<br>
© Syntegon Group.<br>
All rights reserved, also regarding any disposal, exploitation, reproduction, editing, distribution,<br>
as well as in the event of applications for industrial property rights.<br>
*****************************************************************************************************<br>
DESCRIPTION:<br>
XTS gantry: the movers follow up to four products on the IDH infeed (the most downstream mover takes the<br>
first product), then the Z axis lowers all grippers together, the X axes carry the products over the tray<br>
belt, they are put down together and the movers return to their waiting positions.<br>
****************************************************************************************************)
METHOD PRIVATE m_Step : BOOL
VAR
	n_TempI								: INT;
	un_TempIndex						: UINT;
	udn_TempBest						: UDINT;	// [-] product id
	lr_TempBest							: LREAL;	// [mm]
	lr_TempPos							: LREAL;	// [mm]
	lr_TempRz							: LREAL;	// [deg]
	n_TempAssigned						: INT;
	b_TempAllSynced						: BOOL;
	b_TempAnySynced						: BOOL;
	b_TempDone							: BOOL;
	b_TempSynced						: ARRAY[0..3] OF BOOL;
	TempProduct							: ST_VisuProduct;
	TempPose							: ST_VisuPlanarPose;
	TempLatch							: ST_VisuPlanarPose;
END_VAR
(****************************************************************************************************)
(* SEQUENCE                                                                                         *)
(****************************************************************************************************)
CASE n_GantryPhase OF
	n_GANTRY_COLLECT:
		(* Downstream mover first: it takes the most downstream product not yet assigned. *)
		FOR n_TempI := 3 TO 0 BY -1 DO
			IF udn_GantryProduct[n_TempI] = 0 THEN
				udn_TempBest := 0;
				lr_TempBest := -1.0E9;
				FOR un_TempIndex := 1 TO fb_IdhInfeed.m_ProductCount() DO
					fb_IdhInfeed.m_GetProduct(vi_un_Index := un_TempIndex - 1, vo_Product => TempProduct, vo_Pose => TempPose);
					TempPose := fb_IdhInfeed.m_BeltToMcs(vi_Pose := TempPose);
					lr_TempPos := TempPose.fX - lr_GANTRY_X;
					IF TempProduct.eState = E_VisuProductState.DETECTED AND lr_TempPos < lr_GantryPos[n_TempI]
					AND lr_TempPos > -500 AND lr_TempPos > lr_TempBest
					THEN
						udn_TempBest := TempProduct.nId;
						lr_TempBest := lr_TempPos;
					END_IF
				END_FOR
				IF udn_TempBest = 0 THEN
					EXIT;
				END_IF
				fb_IdhInfeed.m_SetProductState(vi_udn_Id := udn_TempBest, vi_e_State := E_VisuProductState.ASSIGNED,
					vi_udn_ClientId := fb_Idh.m_Id(), vi_udn_MoverId := INT_TO_UDINT(n_TempI + 1), vi_udn_FingerId := 0);
				udn_GantryProduct[n_TempI] := udn_TempBest;
			END_IF
		END_FOR
		m_Follow();

		(* Pick once all four are above their products, or at the track end with any of them. *)
		n_TempAssigned := 0;
		b_TempAllSynced := TRUE;
		b_TempAnySynced := FALSE;
		FOR n_TempI := 0 TO 3 DO
			b_TempSynced[n_TempI] := FALSE;
			IF udn_GantryProduct[n_TempI] <> 0 THEN
				n_TempAssigned := n_TempAssigned + 1;
				b_TempSynced[n_TempI] := m_TrackPos(vi_udn_Id := udn_GantryProduct[n_TempI], vo_lr_TrackPos => lr_TempPos,
											vo_lr_Rz => lr_TempRz)
										AND ABS(lr_GantryPos[n_TempI] - lr_TempPos) < 2;
				b_TempAllSynced := b_TempAllSynced AND b_TempSynced[n_TempI];
				b_TempAnySynced := b_TempAnySynced OR b_TempSynced[n_TempI];
			END_IF
		END_FOR
		IF (n_TempAssigned = 4 AND b_TempAllSynced)
		OR (lr_GantryPos[3] >= UINT_TO_LREAL(un_GANTRY_MODULES) * lr_GANTRY_MODULE_LENGTH - 300 AND b_TempAnySynced)
		THEN
			(* Movers not yet above their product give it back. *)
			FOR n_TempI := 0 TO 3 DO
				IF udn_GantryProduct[n_TempI] <> 0 AND NOT b_TempSynced[n_TempI] THEN
					fb_IdhInfeed.m_SetProductState(vi_udn_Id := udn_GantryProduct[n_TempI],
						vi_e_State := E_VisuProductState.DETECTED, vi_udn_ClientId := fb_Idh.m_Id(), vi_udn_MoverId := 0,
						vi_udn_FingerId := 0);
					udn_GantryProduct[n_TempI] := 0;
				END_IF
			END_FOR
			n_GantryPhase := n_GANTRY_PICK_DOWN;
		END_IF

	n_GANTRY_PICK_DOWN:
		m_Follow();
		lr_GantryZ := _FC_DemoApproach(lr_GantryZ, lr_GANTRY_Z_DOWN, lr_GANTRY_Z_SPEED * lr_Dt);
		IF lr_GantryZ = lr_GANTRY_Z_DOWN THEN
			FOR n_TempI := 0 TO 3 DO
				IF udn_GantryProduct[n_TempI] <> 0 THEN
					b_GantryGrip[n_TempI] := TRUE;
					fb_IdhInfeed.m_SetProductState(vi_udn_Id := udn_GantryProduct[n_TempI], vi_e_State := E_VisuProductState.PICKED,
						vi_udn_ClientId := fb_Idh.m_Id(), vi_udn_MoverId := INT_TO_UDINT(n_TempI + 1), vi_udn_FingerId := 1);
				END_IF
			END_FOR
			n_GantryPhase := n_GANTRY_PICK_UP;
		END_IF

	n_GANTRY_PICK_UP:
		lr_GantryZ := _FC_DemoApproach(lr_GantryZ, 0, lr_GANTRY_Z_SPEED * lr_Dt);
		IF lr_GantryZ = 0 THEN
			n_GantryPhase := n_GANTRY_TO_TRAY;
		END_IF

	n_GANTRY_TO_TRAY:
		b_TempDone := TRUE;
		FOR n_TempI := 0 TO 3 DO
			lr_GantryX[n_TempI] := _FC_DemoApproach(lr_GantryX[n_TempI], lr_GANTRY_X_TRAY, lr_GANTRY_X_SPEED * lr_Dt);
			lr_GantryC[n_TempI] := _FC_DemoApproach(lr_GantryC[n_TempI], 0, 180.0 * lr_Dt);
			b_TempDone := b_TempDone AND lr_GantryX[n_TempI] = lr_GANTRY_X_TRAY AND lr_GantryC[n_TempI] = 0;
		END_FOR
		IF b_TempDone THEN
			n_GantryPhase := n_GANTRY_PLACE_DOWN;
		END_IF

	n_GANTRY_PLACE_DOWN:
		lr_GantryZ := _FC_DemoApproach(lr_GantryZ, lr_GANTRY_Z_DOWN, lr_GANTRY_Z_SPEED * lr_Dt);
		IF lr_GantryZ = lr_GANTRY_Z_DOWN THEN
			FOR n_TempI := 0 TO 3 DO
				IF udn_GantryProduct[n_TempI] <> 0 THEN
					(* Put down on the tray: it no longer lies on the infeed. *)
					fb_IdhInfeed.m_RemoveProduct(udn_GantryProduct[n_TempI]);
					(* Turned by -90 deg: gripper at MCS x = track start + position, y = pose y - (X + tool offset). *)
					TempLatch.fX := lr_GANTRY_X + lr_GantryPos[n_TempI];
					TempLatch.fY := lr_GANTRY_Y - (lr_GantryX[n_TempI] + lr_GANTRY_TOOL_X);
					TempLatch.fZ := DEMO_GlobalConst.DEMO_lr_BELT_Z;
					TempLatch.fRz := -90 + lr_GantryC[n_TempI];	// as the cup holds it
					IF fb_IdhTray.m_LatchProduct(vi_udn_Id := DEMO_GlobalVar.DEMO_udn_NextId,
						vi_LatchPose := fb_IdhTray.m_McsToBelt(vi_Pose := TempLatch),
						vi_udn_ProductType := 1, vi_lr_LatchBeltPosition := 0, vi_b_UseLatchBeltPosition := FALSE,
						vi_e_State := E_VisuProductState.PLACED, vi_udn_ClientId := fb_Idh.m_Id())
					THEN
						DEMO_GlobalVar.DEMO_udn_NextId := DEMO_GlobalVar.DEMO_udn_NextId + 1;
					END_IF
					udn_GantryProduct[n_TempI] := 0;
				END_IF
				b_GantryGrip[n_TempI] := FALSE;
			END_FOR
			n_GantryPhase := n_GANTRY_PLACE_UP;
		END_IF

	n_GANTRY_PLACE_UP:
		lr_GantryZ := _FC_DemoApproach(lr_GantryZ, 0, lr_GANTRY_Z_SPEED * lr_Dt);
		IF lr_GantryZ = 0 THEN
			n_GantryPhase := n_GANTRY_RETURN;
		END_IF

	n_GANTRY_RETURN:
		m_Follow();
		b_TempDone := TRUE;
		FOR n_TempI := 0 TO 3 DO
			lr_GantryX[n_TempI] := _FC_DemoApproach(lr_GantryX[n_TempI], lr_GANTRY_X_BELT, lr_GANTRY_X_SPEED * lr_Dt);
			b_TempDone := b_TempDone AND lr_GantryX[n_TempI] = lr_GANTRY_X_BELT AND lr_GantryPos[n_TempI] = lr_GantryWait[n_TempI];
		END_FOR
		IF b_TempDone THEN
			n_GantryPhase := n_GANTRY_COLLECT;
		END_IF
END_CASE


(****************************************************************************************************)
(* REPORT                                                                                           *)
(****************************************************************************************************)
fb_Idh.m_SetZPosition(lr_GantryZ);
fb_Idh.m_SetMoverCount(4);
FOR n_TempI := 0 TO 3 DO
	(* The cup hangs from the flange and turns only about Rz, by the gripper's C. Turned by -90 deg: local (x, y, z)
	   is MCS (gantry x + y, gantry y - x, gantry z + z). *)
	MoverFingers[0].stPose.fX := lr_GANTRY_X + lr_GantryPos[n_TempI];
	MoverFingers[0].stPose.fY := lr_GANTRY_Y - (lr_GantryX[n_TempI] + lr_GANTRY_TOOL_X);
	MoverFingers[0].stPose.fZ := lr_GANTRY_Z + lr_GantryZ + lr_GANTRY_TOOL_Z + DEMO_GlobalConst.DEMO_lr_CUP_HEIGHT;
	MoverFingers[0].stPose.fRx := 0;
	MoverFingers[0].stPose.fRy := 0;
	MoverFingers[0].stPose.fRz := -90 + lr_GantryC[n_TempI];
	MoverFingers[0].bActive := b_GantryGrip[n_TempI];
	(* Demo fault: mover 2 now and then. *)
	fb_Idh.m_SetMover(vi_un_Index := INT_TO_UINT(n_TempI), vi_udn_Id := INT_TO_UDINT(n_TempI + 1),
		vi_lr_Position := lr_GantryPos[n_TempI], vi_lr_X := lr_GantryX[n_TempI], vi_b_GripperActive := b_GantryGrip[n_TempI],
		vi_FingerStates := MoverFingers,
		vi_b_Fault := n_TempI = 1 AND DEMO_GlobalVar.DEMO_lr_FaultPhase >= lr_FAULT_START
					AND DEMO_GlobalVar.DEMO_lr_FaultPhase < lr_FAULT_START + DEMO_GlobalConst.DEMO_lr_FAULT_DURATION,
		vi_str_FaultMessage := 'Vacuum not reached');
END_FOR
m_Step := TRUE;
END_METHOD

(****************************************************************************************************<br>
© Syntegon Group.<br>
All rights reserved, also regarding any disposal, exploitation, reproduction, editing, distribution,<br>
as well as in the event of applications for industrial property rights.<br>
*****************************************************************************************************<br>
DESCRIPTION:<br>
Position of a product on the IDH infeed along the gantry track (MCS x - gantry x) and its rotation.<br>
FALSE if the product is no longer in the register.<br>
****************************************************************************************************)
METHOD PRIVATE m_TrackPos : BOOL
VAR_INPUT
	vi_udn_Id							: UDINT;	// [-] product id
END_VAR
VAR_OUTPUT
	vo_lr_TrackPos						: LREAL;	// [mm]
	vo_lr_Rz							: LREAL;	// [deg]
END_VAR
VAR
	n_TempIndex							: INT;
	TempProduct							: ST_VisuProduct;
	TempPose							: ST_VisuPlanarPose;
END_VAR
n_TempIndex := fb_IdhInfeed.m_FindProduct(vi_udn_Id);
m_TrackPos := n_TempIndex >= 0;
IF m_TrackPos THEN
	fb_IdhInfeed.m_GetProduct(vi_un_Index := INT_TO_UINT(n_TempIndex), vo_Product => TempProduct, vo_Pose => TempPose);
	TempPose := fb_IdhInfeed.m_BeltToMcs(vi_Pose := TempPose);
	vo_lr_TrackPos := TempPose.fX - lr_GANTRY_X;
	vo_lr_Rz := TempPose.fRz;
END_IF
END_METHOD

END_PROGRAM

// ---- POUs/P_VisuDemoCartesian.TcPOU
(****************************************************************************************************<br>
© Syntegon Group.<br>
All rights reserved, also regarding any disposal, exploitation, reproduction, editing, distribution,<br>
as well as in the event of applications for industrial property rights.<br>
*****************************************************************************************************<br>
DESCRIPTION:<br>
DEMO ONLY: Cartesian application (Y = 6500..7300). A Cartesian robot picks products from the Cartesian infeed,<br>
turns them by C = -90 deg, tilts them by A while lowering and places them onto the Cartesian outfeed, every second<br>
one on top of the one it put down before (following it along the belt). Its gripper<br>
is a cup in the middle with two jaws beside it. Called by P_VisuDemo.<br>
****************************************************************************************************)
PROGRAM P_VisuDemoCartesian
VAR
	fb_CartInfeed						: _FB_VisuConveyor;
	fb_CartOutfeed						: _FB_VisuConveyor;
	fb_Cartesian						: _FB_VisuCartesian;

	(* Conveyors *)
	lr_Dt								: LREAL;	// [s] cycle time
	udn_Seed							: UDINT := 45678;	// [-] pseudo random generator state
	lr_InfeedPosition					: LREAL;	// [mm] belt position of the Cartesian infeed
	lr_OutfeedPosition					: LREAL;	// [mm] belt position of the Cartesian outfeed
	lr_SinceSpawn						: LREAL;	// [s] since the last product
	BeltPose							: ST_VisuPose;
	LatchPose							: ST_VisuPlanarPose;
	CartPose							: ST_VisuPose;

	(* Cartesian robot: axis actual values, start above the infeed *)
	n_CartPhase							: INT;
	lr_CartX							: LREAL := 900;	// [mm]
	lr_CartY							: LREAL := 200;	// [mm]
	lr_CartZ							: LREAL := -200;	// [mm]
	lr_CartC							: LREAL;	// [deg]
	lr_CartA							: LREAL;	// [deg]
	lr_CartPickC						: LREAL;	// [deg] C that turns the gripper onto the current product
	lr_CartJaw							: LREAL := 120;	// [mm] jaw distance from the cup along the gripper's X
	b_CartGrip							: BOOL;
	udn_CartProduct						: UDINT;	// [-] product id on the Cartesian infeed
	udn_CartStackBase					: UDINT;	// [-] product on the outfeed the next one is stacked on, 0 = the next one becomes it
	b_CartStacking						: BOOL;	// the product carried now goes onto udn_CartStackBase
END_VAR
VAR CONSTANT
	(* Robot turned by -90 deg: X axis across the belts towards MCS -Y (outfeed under X = 100, infeed under
	   X = 900), Y axis along MCS +X from X = 1000. *)
	lr_CART_INFEED_Y					: LREAL := 6500;	// [mm]
	lr_CART_OUTFEED_Y					: LREAL := 7300;	// [mm]
	lr_CART_BELT_LENGTH					: LREAL := 3000;	// [mm]
	lr_CART_BELT_SPEED					: LREAL := 150;	// [mm/s]
	lr_CART_SPAWN_INTERVAL				: LREAL := 2.5;	// [s]
	lr_CART_X							: LREAL := 1000;	// [mm]
	lr_CART_Y							: LREAL := 7400;	// [mm]
	lr_CART_Z							: LREAL := 1540;	// [mm] Z = -550 puts the cup's grip point (A = 0) on the product top
	lr_CART_TOOL_LENGTH					: LREAL := 150;	// [mm] flange to the cup's grip point
	lr_CART_CUP_HEIGHT					: LREAL := 40;	// [mm]
	lr_CART_JAW_DIAMETER				: LREAL := 20;	// [mm]
	lr_CART_JAW_HEIGHT					: LREAL := 120;	// [mm]
	lr_CART_JAW_TOP						: LREAL := 60;	// [mm] jaw tops below the flange
	lr_CART_JAW_OPEN					: LREAL := 120;	// [mm]
	lr_CART_JAW_CLOSED					: LREAL := 70;	// [mm] closed on a 120 mm product
	lr_CART_JAW_SPEED					: LREAL := 300;	// [mm/s]
	lr_CART_RAIL_HEIGHT					: LREAL := 1200;	// [mm]
	lr_CART_X_OUTFEED					: LREAL := 100;	// [mm]
	lr_CART_X_INFEED					: LREAL := 900;	// [mm]
	lr_CART_Y_HOME						: LREAL := 200;	// [mm]
	lr_CART_Y_STACK_BASE				: LREAL := 300;	// [mm] a product the next one is stacked on is put down here
	lr_CART_Y_STACK_MAX				: LREAL := 900;	// [mm] beyond this no stacking: the product below would leave the reach
	lr_CART_Z_PICK						: LREAL := -550;	// [mm]
	lr_CART_Z_TRAVEL					: LREAL := -200;	// [mm]
	lr_CART_TILT						: LREAL := 20;	// [deg] A while lowering
	lr_CART_TURN						: LREAL := -90;	// [deg] C between pick and place
	lr_CART_XY_SPEED					: LREAL := 1500;	// [mm/s]
	lr_CART_Z_SPEED						: LREAL := 800;	// [mm/s]
	lr_CART_C_SPEED						: LREAL := 180;	// [deg/s]
	lr_CART_A_SPEED						: LREAL := 60;	// [deg/s]
	n_CART_IDLE							: INT := 0;
	n_CART_DESCEND						: INT := 1;
	n_CART_LIFT							: INT := 2;
	n_CART_TRANSFER						: INT := 3;
	n_CART_LOWER						: INT := 4;
	n_CART_STRAIGHTEN					: INT := 5;
	n_CART_RELEASE						: INT := 6;
	n_CART_RISE							: INT := 7;
END_VAR

lr_Dt := DEMO_GlobalVar.DEMO_lr_Dt;


(****************************************************************************************************)
(* REGISTRATION (idempotent, every cycle)                                                           *)
(****************************************************************************************************)
fb_CartInfeed.m_Register(vio_Manifest := GVL_Visu.stManifest, vi_udn_Id := 8, vi_str_Name := 'Cartesian infeed');
fb_CartOutfeed.m_Register(vio_Manifest := GVL_Visu.stManifest, vi_udn_Id := 9, vi_str_Name := 'Cartesian outfeed');
fb_Cartesian.m_Register(vio_Manifest := GVL_Visu.stManifest, vi_udn_Id := 40, vi_str_Name := 'Cartesian');


(****************************************************************************************************)
(* CONVEYORS (configuration idempotent, every cycle)                                                *)
(****************************************************************************************************)
BeltPose.fX := 0;
BeltPose.fY := lr_CART_INFEED_Y;
BeltPose.fZ := DEMO_GlobalConst.DEMO_lr_BELT_Z;
fb_CartInfeed.m_SetPose(vi_Pose := BeltPose);
fb_CartInfeed.m_Configure(vi_lr_Length := lr_CART_BELT_LENGTH,
	vi_lr_Width := DEMO_GlobalConst.DEMO_lr_BELT_WIDTH);
BeltPose.fY := lr_CART_OUTFEED_Y;
fb_CartOutfeed.m_SetPose(vi_Pose := BeltPose);
fb_CartOutfeed.m_Configure(vi_lr_Length := lr_CART_BELT_LENGTH,
	vi_lr_Width := DEMO_GlobalConst.DEMO_lr_BELT_WIDTH);
(* The infeed's belt coordinates count from the robot's Y = 0, 1000 mm behind the belt start. *)
fb_CartInfeed.m_SetOriginShift(vi_lr_X := lr_CART_X, vi_lr_Y := 0, vi_lr_Z := 0);
fb_CartInfeed.m_SetProductType(vi_udn_Id := 1, vi_lr_Length := DEMO_GlobalConst.DEMO_lr_PRODUCT_LENGTH,
	vi_lr_Width := DEMO_GlobalConst.DEMO_lr_PRODUCT_WIDTH, vi_lr_Height := DEMO_GlobalConst.DEMO_lr_PRODUCT_HEIGHT,
	vi_e_Shape := E_VisuProductShape.BOX, vi_lr_CornerRadius := 0);
fb_CartOutfeed.m_SetProductType(vi_udn_Id := 1, vi_lr_Length := DEMO_GlobalConst.DEMO_lr_PRODUCT_LENGTH,
	vi_lr_Width := DEMO_GlobalConst.DEMO_lr_PRODUCT_WIDTH, vi_lr_Height := DEMO_GlobalConst.DEMO_lr_PRODUCT_HEIGHT,
	vi_e_Shape := E_VisuProductShape.BOX, vi_lr_CornerRadius := 0);

(* Belt travel *)
lr_InfeedPosition := lr_InfeedPosition + lr_CART_BELT_SPEED * lr_Dt;
lr_OutfeedPosition := lr_OutfeedPosition + lr_CART_BELT_SPEED * lr_Dt;
fb_CartInfeed.m_SetBeltPosition(lr_InfeedPosition);
fb_CartOutfeed.m_SetBeltPosition(lr_OutfeedPosition);


(****************************************************************************************************)
(* PRODUCT INFEED: regular gaps, products turned                                                    *)
(****************************************************************************************************)
lr_SinceSpawn := lr_SinceSpawn + lr_Dt;
IF lr_SinceSpawn >= lr_CART_SPAWN_INTERVAL THEN
	lr_SinceSpawn := 0;
	udn_Seed := udn_Seed * 1103515245 + 12345;
	LatchPose.fX := 100;
	LatchPose.fY := lr_CART_INFEED_Y;
	LatchPose.fZ := DEMO_GlobalConst.DEMO_lr_BELT_Z;
	LatchPose.fRz := (UDINT_TO_LREAL((udn_Seed / 1000) MOD 1000) / 1000.0 - 0.5) * 60.0;
	IF fb_CartInfeed.m_LatchProduct(vi_udn_Id := DEMO_GlobalVar.DEMO_udn_NextId,
		vi_LatchPose := fb_CartInfeed.m_McsToBelt(vi_Pose := LatchPose),
		vi_udn_ProductType := 1, vi_lr_LatchBeltPosition := 0, vi_b_UseLatchBeltPosition := FALSE,
		vi_e_State := E_VisuProductState.DETECTED, vi_udn_ClientId := 0)
	THEN
		DEMO_GlobalVar.DEMO_udn_NextId := DEMO_GlobalVar.DEMO_udn_NextId + 1;
	END_IF
END_IF


(****************************************************************************************************)
(* CARTESIAN ROBOT                                                                                  *)
(****************************************************************************************************)
CartPose.fX := lr_CART_X;
CartPose.fY := lr_CART_Y;
CartPose.fZ := lr_CART_Z;
CartPose.fRz := -90;
fb_Cartesian.m_SetPose(vi_Pose := CartPose);
fb_Cartesian.m_Configure(vi_lr_XMin := 0, vi_lr_XMax := 1200, vi_lr_YMin := 0, vi_lr_YMax := 1000,
	vi_lr_ZMin := -600, vi_lr_ZMax := 0, vi_lr_RailHeight := lr_CART_RAIL_HEIGHT);
(* Limit area in the robot frame (flange coordinates): X only up to the infeed, Z not into the top 100 mm. *)
fb_Cartesian.m_SetLimitArea(vi_lr_XMin := 0, vi_lr_XMax := 1000, vi_lr_YMin := 0, vi_lr_YMax := 1000,
	vi_lr_ZMin := -600, vi_lr_ZMax := -100);
(* Around the flange and the gripper below it. *)
fb_Cartesian.m_SetTcpLimitArea(vi_lr_XMin := -80, vi_lr_XMax := 80, vi_lr_YMin := -80, vi_lr_YMax := 80,
	vi_lr_ZMin := -50, vi_lr_ZMax := 20);
(* A cup in the middle carries the product, two jaws close beside it. *)
fb_Cartesian.m_SetFinger(vi_un_Finger := 1, vi_lr_Diameter := DEMO_GlobalConst.DEMO_lr_CUP_DIAMETER,
	vi_lr_Height := lr_CART_CUP_HEIGHT);
fb_Cartesian.m_SetFinger(vi_un_Finger := 2, vi_lr_Diameter := lr_CART_JAW_DIAMETER, vi_lr_Height := lr_CART_JAW_HEIGHT);
fb_Cartesian.m_SetFinger(vi_un_Finger := 3, vi_lr_Diameter := lr_CART_JAW_DIAMETER, vi_lr_Height := lr_CART_JAW_HEIGHT);
fb_Cartesian.m_SetZone(vi_un_Zone := 1, vi_udn_ConveyorId := fb_CartInfeed.m_Id(),
	vi_lr_Start := 0, vi_lr_End := 1000, vi_lr_AllocationOffset := 0, vi_lr_CcsOffset := 0,
	vi_lr_StartY := 0, vi_lr_EndY := 0);
fb_Cartesian.m_SetZone(vi_un_Zone := 2, vi_udn_ConveyorId := fb_CartOutfeed.m_Id(),
	vi_lr_Start := lr_CART_X + lr_CART_Y_STACK_BASE - 100, vi_lr_End := lr_CART_X + lr_CART_Y_STACK_MAX + 100,
	vi_lr_AllocationOffset := 0, vi_lr_CcsOffset := lr_CART_X + (lr_CART_Y_STACK_BASE + lr_CART_Y_STACK_MAX) / 2,
	vi_lr_StartY := 0, vi_lr_EndY := 0);
m_Step();
fb_Cartesian.m_SetAxes(vi_lr_X := lr_CartX, vi_lr_Y := lr_CartY, vi_lr_Z := lr_CartZ, vi_b_GripperActive := b_CartGrip);

(* C and A turn and tilt the gripper below the flange; they show only through the finger poses. *)
lr_CartJaw := _FC_DemoApproach(lr_CartJaw, SEL(b_CartGrip, lr_CART_JAW_OPEN, lr_CART_JAW_CLOSED), lr_CART_JAW_SPEED * lr_Dt);
fb_Cartesian.m_SetFingerState(vi_un_Finger := 1,
	vi_Pose := m_Finger(vi_lr_OffsetX := 0, vi_lr_OffsetZ := -(lr_CART_TOOL_LENGTH - lr_CART_CUP_HEIGHT)),
	vi_b_Active := b_CartGrip);
fb_Cartesian.m_SetFingerState(vi_un_Finger := 2,
	vi_Pose := m_Finger(vi_lr_OffsetX := lr_CartJaw, vi_lr_OffsetZ := -lr_CART_JAW_TOP),
	vi_b_Active := b_CartGrip);
fb_Cartesian.m_SetFingerState(vi_un_Finger := 3,
	vi_Pose := m_Finger(vi_lr_OffsetX := -lr_CartJaw, vi_lr_OffsetZ := -lr_CART_JAW_TOP),
	vi_b_Active := b_CartGrip);


(****************************************************************************************************)
(* HOUSEKEEPING                                                                                     *)
(****************************************************************************************************)
fb_CartInfeed.m_RemoveProductsBeyond(lr_CART_BELT_LENGTH + DEMO_GlobalConst.DEMO_lr_REMOVE_BEYOND_END);
fb_CartOutfeed.m_RemoveProductsBeyond(lr_CART_BELT_LENGTH + DEMO_GlobalConst.DEMO_lr_REMOVE_BEYOND_END);

(****************************************************************************************************<br>
© Syntegon Group.<br>
All rights reserved, also regarding any disposal, exploitation, reproduction, editing, distribution,<br>
as well as in the event of applications for industrial property rights.<br>
*****************************************************************************************************<br>
DESCRIPTION:<br>
Pose of a Cartesian gripper finger, absolute in the MCS: the finger sits at (vi_lr_OffsetX, 0, vi_lr_OffsetZ) in<br>
the gripper, which is turned by C about Z and tilted by A about its own X below the flange. The robot is<br>
turned by -90 deg: local (x, y, z) is MCS (lr_CART_X + y, lr_CART_Y - x, lr_CART_Z + z).<br>
****************************************************************************************************)
METHOD PRIVATE m_Finger : ST_VisuPose
VAR_INPUT
	vi_lr_OffsetX						: LREAL;	// [mm] along the gripper's X
	vi_lr_OffsetZ						: LREAL;	// [mm] below the flange: negative
END_VAR
VAR
	lr_TempA							: LREAL;	// [rad]
	lr_TempC							: LREAL;	// [rad]
	lr_TempVx							: LREAL;	// [mm] offset in the robot frame
	lr_TempVy							: LREAL;	// [mm]
	lr_TempVz							: LREAL;	// [mm]
END_VAR
lr_TempA := lr_CartA * VISU_GlobalConst.VISU_lr_DEG_TO_RAD;
lr_TempC := lr_CartC * VISU_GlobalConst.VISU_lr_DEG_TO_RAD;
(* Rz(C) * Rx(A) * (x, 0, z) *)
lr_TempVx := vi_lr_OffsetX * COS(lr_TempC) + vi_lr_OffsetZ * SIN(lr_TempA) * SIN(lr_TempC);
lr_TempVy := vi_lr_OffsetX * SIN(lr_TempC) - vi_lr_OffsetZ * SIN(lr_TempA) * COS(lr_TempC);
lr_TempVz := vi_lr_OffsetZ * COS(lr_TempA);
m_Finger.fX := lr_CART_X + (lr_CartY + lr_TempVy);
m_Finger.fY := lr_CART_Y - (lr_CartX + lr_TempVx);
m_Finger.fZ := lr_CART_Z + (lr_CartZ + lr_TempVz);
m_Finger.fRx := lr_CartA;
m_Finger.fRy := 0;
m_Finger.fRz := -90 + lr_CartC;
END_METHOD

(****************************************************************************************************<br>
© Syntegon Group.<br>
All rights reserved, also regarding any disposal, exploitation, reproduction, editing, distribution,<br>
as well as in the event of applications for industrial property rights.<br>
*****************************************************************************************************<br>
DESCRIPTION:<br>
Moves the Cartesian robot's axes one cycle towards the goal, each with its own speed. TRUE once all are there.<br>
****************************************************************************************************)
METHOD PRIVATE m_Move : BOOL
VAR_INPUT
	vi_lr_X								: LREAL;	// [mm]
	vi_lr_Y								: LREAL;	// [mm]
	vi_lr_Z								: LREAL;	// [mm]
	vi_lr_C								: LREAL;	// [deg]
	vi_lr_A								: LREAL;	// [deg]
END_VAR
lr_CartX := _FC_DemoApproach(lr_CartX, vi_lr_X, lr_CART_XY_SPEED * lr_Dt);
lr_CartY := _FC_DemoApproach(lr_CartY, vi_lr_Y, lr_CART_XY_SPEED * lr_Dt);
lr_CartZ := _FC_DemoApproach(lr_CartZ, vi_lr_Z, lr_CART_Z_SPEED * lr_Dt);
lr_CartC := _FC_DemoApproach(lr_CartC, vi_lr_C, lr_CART_C_SPEED * lr_Dt);
lr_CartA := _FC_DemoApproach(lr_CartA, vi_lr_A, lr_CART_A_SPEED * lr_Dt);
(* _FC_DemoApproach lands exactly on the goal, so equality is safe. *)
m_Move := lr_CartX = vi_lr_X AND lr_CartY = vi_lr_Y AND lr_CartZ = vi_lr_Z AND lr_CartC = vi_lr_C AND lr_CartA = vi_lr_A;
END_METHOD

(****************************************************************************************************<br>
© Syntegon Group.<br>
All rights reserved, also regarding any disposal, exploitation, reproduction, editing, distribution,<br>
as well as in the event of applications for industrial property rights.<br>
*****************************************************************************************************<br>
DESCRIPTION:<br>
Cartesian robot: follows a product on the Cartesian infeed in Y with the gripper turned onto it (C), picks<br>
it, carries it across to the outfeed while turning it by a further -90 deg, tilts it by A while lowering,<br>
straightens it and places it. Every second product goes on top of the one put down before, following it along<br>
the outfeed, as long as that one is in reach; otherwise it is put down at lr_CART_Y_STACK_BASE and the next one<br>
is stacked on it.<br>
****************************************************************************************************)
METHOD PRIVATE m_Step : BOOL
VAR
	n_TempFound							: INT;
	un_TempScan							: UINT;
	b_TempHave							: BOOL;
	lr_TempProductY						: LREAL;	// [mm] robot Y of the current product: its MCS x relative to the robot origin
	TempProduct							: ST_VisuProduct;
	TempProductPose						: ST_VisuPlanarPose;
	TempPlacePose						: ST_VisuPlanarPose;
	TempStackProduct					: ST_VisuProduct;
	TempStackPose						: ST_VisuPlanarPose;
	n_TempStackIdx						: INT;
	b_TempStackFound					: BOOL;
	lr_TempStackY						: LREAL;	// [mm] robot Y of the product to stack on
	lr_TempPlaceY						: LREAL;	// [mm] robot Y to put the product down at
	lr_TempPlaceZ						: LREAL;	// [mm] robot Z to put it down at: one product higher when stacking
	udn_TempPlacedId					: UDINT;
END_VAR
(* Current product *)
b_TempHave := FALSE;
IF udn_CartProduct <> 0 THEN
	n_TempFound := fb_CartInfeed.m_FindProduct(udn_CartProduct);
	IF n_TempFound >= 0 THEN
		b_TempHave := fb_CartInfeed.m_GetProduct(vi_un_Index := INT_TO_UINT(n_TempFound), vo_Product => TempProduct,
			vo_Pose => TempProductPose);
		TempProductPose := fb_CartInfeed.m_BeltToMcs(vi_Pose := TempProductPose);
		lr_TempProductY := TempProductPose.fX - lr_CART_X;
	END_IF
END_IF

(* Product to stack on, while it travels on the outfeed *)
b_TempStackFound := FALSE;
IF udn_CartStackBase <> 0 THEN
	n_TempStackIdx := fb_CartOutfeed.m_FindProduct(udn_CartStackBase);
	IF n_TempStackIdx >= 0 THEN
		fb_CartOutfeed.m_GetProduct(vi_un_Index := INT_TO_UINT(n_TempStackIdx), vo_Product => TempStackProduct,
			vo_Pose => TempStackPose);
		TempStackPose := fb_CartOutfeed.m_BeltToMcs(vi_Pose := TempStackPose);
		lr_TempStackY := TempStackPose.fX - lr_CART_X;
		b_TempStackFound := TRUE;
	END_IF
END_IF
IF NOT b_TempStackFound THEN
	b_CartStacking := FALSE;
END_IF
lr_TempPlaceY := SEL(b_CartStacking, lr_CART_Y_STACK_BASE, lr_TempStackY);
lr_TempPlaceZ := lr_CART_Z_PICK + SEL(b_CartStacking, 0, DEMO_GlobalConst.DEMO_lr_PRODUCT_HEIGHT);

(* Sequence *)
CASE n_CartPhase OF
	n_CART_IDLE:
		un_TempScan := 0;
		WHILE udn_CartProduct = 0 AND un_TempScan < fb_CartInfeed.m_ProductCount() DO
			fb_CartInfeed.m_GetProduct(vi_un_Index := un_TempScan, vo_Product => TempProduct, vo_Pose => TempProductPose);
			TempProductPose := fb_CartInfeed.m_BeltToMcs(vi_Pose := TempProductPose);
			IF TempProduct.eState = E_VisuProductState.DETECTED
			AND TempProductPose.fX - lr_CART_X >= 100
			AND TempProductPose.fX - lr_CART_X <= 600
			THEN
				fb_CartInfeed.m_SetProductState(vi_udn_Id := TempProduct.nId, vi_e_State := E_VisuProductState.ASSIGNED,
					vi_udn_ClientId := fb_Cartesian.m_Id(), vi_udn_MoverId := 0, vi_udn_FingerId := 0);
				udn_CartProduct := TempProduct.nId;
				(* The gripper's +X in the MCS is pose rz (-90 deg) + C. *)
				lr_CartPickC := TempProductPose.fRz + 90;
				n_CartPhase := n_CART_DESCEND;
			END_IF
			un_TempScan := un_TempScan + 1;
		END_WHILE
		IF udn_CartProduct = 0 THEN
			m_Move(vi_lr_X := lr_CART_X_INFEED, vi_lr_Y := lr_CART_Y_HOME, vi_lr_Z := lr_CART_Z_TRAVEL, vi_lr_C := 0,
				vi_lr_A := 0);
		END_IF

	n_CART_DESCEND:
		IF NOT b_TempHave THEN
			udn_CartProduct := 0;
			n_CartPhase := n_CART_RISE;
		ELSIF lr_TempProductY > 1000 THEN
			(* Out of reach: hand it back, it will be missed. *)
			fb_CartInfeed.m_SetProductState(vi_udn_Id := udn_CartProduct, vi_e_State := E_VisuProductState.DETECTED,
				vi_udn_ClientId := fb_Cartesian.m_Id(), vi_udn_MoverId := 0, vi_udn_FingerId := 0);
			udn_CartProduct := 0;
			n_CartPhase := n_CART_RISE;
		ELSIF m_Move(vi_lr_X := lr_CART_X_INFEED, vi_lr_Y := lr_TempProductY, vi_lr_Z := lr_CartZ,
			vi_lr_C := lr_CartPickC, vi_lr_A := 0)
		THEN
			(* Lowers only once above the product with the gripper turned onto it. *)
			IF m_Move(vi_lr_X := lr_CART_X_INFEED, vi_lr_Y := lr_TempProductY, vi_lr_Z := lr_CART_Z_PICK,
				vi_lr_C := lr_CartPickC, vi_lr_A := 0)
			THEN
				fb_CartInfeed.m_SetProductState(vi_udn_Id := udn_CartProduct, vi_e_State := E_VisuProductState.PICKED,
					vi_udn_ClientId := fb_Cartesian.m_Id(), vi_udn_MoverId := 0, vi_udn_FingerId := 1);
				b_CartGrip := TRUE;
				n_CartPhase := n_CART_LIFT;
			END_IF
		END_IF

	n_CART_LIFT:
		IF m_Move(vi_lr_X := lr_CartX, vi_lr_Y := lr_CartY, vi_lr_Z := lr_CART_Z_TRAVEL, vi_lr_C := lr_CartC,
			vi_lr_A := lr_CartA)
		THEN
			n_CartPhase := n_CART_TRANSFER;
		END_IF

	n_CART_TRANSFER:
		(* Every second product goes onto the one put down before, as long as that one is in reach. *)
		b_CartStacking := b_TempStackFound AND lr_TempStackY <= lr_CART_Y_STACK_MAX;
		IF NOT b_CartStacking THEN
			udn_CartStackBase := 0;
		END_IF
		lr_TempPlaceY := SEL(b_CartStacking, lr_CART_Y_STACK_BASE, lr_TempStackY);
		lr_TempPlaceZ := lr_CART_Z_PICK + SEL(b_CartStacking, 0, DEMO_GlobalConst.DEMO_lr_PRODUCT_HEIGHT);
		IF m_Move(vi_lr_X := lr_CART_X_OUTFEED, vi_lr_Y := lr_TempPlaceY, vi_lr_Z := lr_CART_Z_TRAVEL,
			vi_lr_C := lr_CartPickC + lr_CART_TURN, vi_lr_A := 0)
		THEN
			n_CartPhase := n_CART_LOWER;
		END_IF

	n_CART_LOWER:
		IF m_Move(vi_lr_X := lr_CartX, vi_lr_Y := lr_TempPlaceY, vi_lr_Z := lr_TempPlaceZ, vi_lr_C := lr_CartC,
			vi_lr_A := lr_CART_TILT)
		THEN
			n_CartPhase := n_CART_STRAIGHTEN;
		END_IF

	n_CART_STRAIGHTEN:
		IF m_Move(vi_lr_X := lr_CartX, vi_lr_Y := lr_TempPlaceY, vi_lr_Z := lr_CartZ, vi_lr_C := lr_CartC, vi_lr_A := 0) THEN
			n_CartPhase := n_CART_RELEASE;
		END_IF

	n_CART_RELEASE:
		(* Put down on the outfeed: it no longer lies on the infeed. *)
		fb_CartInfeed.m_RemoveProduct(udn_CartProduct);
		(* Turned by -90 deg: the cup (A = 0) is at MCS x = origin + Y, y = origin - X; the product keeps the turn. *)
		TempPlacePose.fX := lr_CART_X + lr_CartY;
		TempPlacePose.fY := lr_CART_Y - lr_CartX;
		(* A stacked product lies one product height above the belt. *)
		TempPlacePose.fZ := DEMO_GlobalConst.DEMO_lr_BELT_Z + SEL(b_CartStacking, 0, DEMO_GlobalConst.DEMO_lr_PRODUCT_HEIGHT);
		TempPlacePose.fRz := -90 + lr_CartC;
		udn_TempPlacedId := DEMO_GlobalVar.DEMO_udn_NextId;
		IF fb_CartOutfeed.m_LatchProduct(vi_udn_Id := DEMO_GlobalVar.DEMO_udn_NextId,
			vi_LatchPose := fb_CartOutfeed.m_McsToBelt(vi_Pose := TempPlacePose),
			vi_udn_ProductType := 1, vi_lr_LatchBeltPosition := 0, vi_b_UseLatchBeltPosition := FALSE,
			vi_e_State := E_VisuProductState.PLACED, vi_udn_ClientId := fb_Cartesian.m_Id())
		THEN
			DEMO_GlobalVar.DEMO_udn_NextId := DEMO_GlobalVar.DEMO_udn_NextId + 1;
		END_IF
		(* The next product goes onto this one, unless this one is already on top of another. *)
		IF b_CartStacking THEN
			udn_CartStackBase := 0;
		ELSE
			udn_CartStackBase := udn_TempPlacedId;
		END_IF
		b_CartStacking := FALSE;
		udn_CartProduct := 0;
		b_CartGrip := FALSE;
		n_CartPhase := n_CART_RISE;

	n_CART_RISE:
		IF m_Move(vi_lr_X := lr_CartX, vi_lr_Y := lr_CartY, vi_lr_Z := lr_CART_Z_TRAVEL, vi_lr_C := lr_CartC,
			vi_lr_A := lr_CartA)
		THEN
			n_CartPhase := n_CART_IDLE;
		END_IF
END_CASE
m_Step := TRUE;
END_METHOD

END_PROGRAM

// ---- POUs/P_VisuDemoCartesianAxes.TcPOU
(****************************************************************************************************<br>
© Syntegon Group.<br>
All rights reserved, also regarding any disposal, exploitation, reproduction, editing, distribution,<br>
as well as in the event of applications for industrial property rights.<br>
*****************************************************************************************************<br>
DESCRIPTION:<br>
DEMO ONLY: Cartesian robots with two axes beside the Cartesian application (X = 4000), moving without<br>
products (m_SetKinematics):<br>
- Cartesian X-Z (Y = 6500): no Y axis, a fixed beam along X; it goes back and forth and dips.<br>
- Cartesian X-Y (Y = 7000..7800): no Z axis, the flange stays at Z min; it runs an ellipse.<br>
Called by P_VisuDemo.<br>
****************************************************************************************************)
PROGRAM P_VisuDemoCartesianAxes
VAR
	fb_CartXz							: _FB_VisuCartesian;
	fb_CartXy							: _FB_VisuCartesian;
	lr_Time								: LREAL;	// [s] since start, wraps with the common period
	lr_AngleXz							: LREAL;	// [rad]
	lr_AngleXy							: LREAL;	// [rad]
	RobotPose							: ST_VisuPose;
END_VAR
VAR CONSTANT
	lr_TWO_PI							: LREAL := 6.283185307179586;	// [-]
	lr_CART_AXES_X						: LREAL := 4000;	// [mm] MCS x of both robots' axis origin
	lr_CART_AXES_Z						: LREAL := 1500;	// [mm] MCS z of both robots' axis origin
	lr_CART_XZ_Y						: LREAL := 6500;	// [mm] MCS y of the X-Z robot
	lr_CART_XY_Y						: LREAL := 7000;	// [mm] MCS y of the X-Y robot's Y = 0
	lr_CART_AXES_RAIL_HEIGHT			: LREAL := 800;	// [mm]
	lr_CART_XZ_PERIOD					: LREAL := 6;	// [s]
	lr_CART_XY_PERIOD					: LREAL := 8;	// [s]
	lr_CART_AXES_WRAP					: LREAL := 24;	// [s] common multiple of both periods
END_VAR

(****************************************************************************************************)
(* REGISTRATION AND CONFIGURATION (idempotent, every cycle)                                         *)
(****************************************************************************************************)
fb_CartXz.m_Register(vio_Manifest := GVL_Visu.stManifest, vi_udn_Id := 41, vi_str_Name := 'Cartesian X-Z');
fb_CartXy.m_Register(vio_Manifest := GVL_Visu.stManifest, vi_udn_Id := 42, vi_str_Name := 'Cartesian X-Y');

RobotPose.fX := lr_CART_AXES_X;
RobotPose.fY := lr_CART_XZ_Y;
RobotPose.fZ := lr_CART_AXES_Z;
(* No Y axis: the Y stroke is ignored, a fixed beam along X carries the carriage. *)
fb_CartXz.m_SetPose(vi_Pose := RobotPose);
fb_CartXz.m_Configure(vi_lr_XMin := 0, vi_lr_XMax := 1200, vi_lr_YMin := 0, vi_lr_YMax := 0,
	vi_lr_ZMin := -600, vi_lr_ZMax := 0, vi_lr_RailHeight := lr_CART_AXES_RAIL_HEIGHT);
fb_CartXz.m_SetKinematics(vi_e_Axes := E_VisuCartesianAxes.XZ);

RobotPose.fY := lr_CART_XY_Y;
(* No Z axis: Z max is ignored, the flange stays at Z min. *)
fb_CartXy.m_SetPose(vi_Pose := RobotPose);
fb_CartXy.m_Configure(vi_lr_XMin := 0, vi_lr_XMax := 1200, vi_lr_YMin := 0, vi_lr_YMax := 800,
	vi_lr_ZMin := -500, vi_lr_ZMax := -500, vi_lr_RailHeight := lr_CART_AXES_RAIL_HEIGHT);
fb_CartXy.m_SetKinematics(vi_e_Axes := E_VisuCartesianAxes.XY);


(****************************************************************************************************)
(* MOTION                                                                                           *)
(****************************************************************************************************)
lr_Time := lr_Time + DEMO_GlobalVar.DEMO_lr_Dt;
IF lr_Time >= lr_CART_AXES_WRAP THEN
	lr_Time := lr_Time - lr_CART_AXES_WRAP;
END_IF
lr_AngleXz := lr_TWO_PI * lr_Time / lr_CART_XZ_PERIOD;
lr_AngleXy := lr_TWO_PI * lr_Time / lr_CART_XY_PERIOD;

(* Y and Z of the missing axes are ignored by the visualisation; report 0. *)
fb_CartXz.m_SetAxes(vi_lr_X := 600 - 500 * COS(lr_AngleXz), vi_lr_Y := 0,
	vi_lr_Z := -300 - 250 * COS(2 * lr_AngleXz), vi_b_GripperActive := FALSE);
fb_CartXy.m_SetAxes(vi_lr_X := 600 + 450 * COS(lr_AngleXy), vi_lr_Y := 400 + 300 * SIN(lr_AngleXy),
	vi_lr_Z := 0, vi_b_GripperActive := FALSE);

END_PROGRAM

// ---- POUs/P_VisuDemoSpacing.TcPOU
(****************************************************************************************************<br>
© Syntegon Group.<br>
All rights reserved, also regarding any disposal, exploitation, reproduction, editing, distribution,<br>
as well as in the event of applications for industrial property rights.<br>
*****************************************************************************************************<br>
DESCRIPTION:<br>
DEMO ONLY: Spacing application (Y = 9000). An XTS loop under one belt takes over products arriving with random<br>
gaps and hands them back to the belt with a constant pitch. The pushed product stays on the belt (moved with<br>
m_MoveProduct), so no placeholder appears. Called by P_VisuDemo.<br>
****************************************************************************************************)
PROGRAM P_VisuDemoSpacing
VAR
	fb_SpcBelt							: _FB_VisuConveyor;
	fb_Spc								: _FB_VisuXtsLoop;

	(* Conveyor *)
	lr_Dt								: LREAL;	// [s] cycle time
	udn_Seed							: UDINT := 56789;	// [-] pseudo random generator state
	lr_SpcBeltPosition					: LREAL;	// [mm]
	lr_SpcSinceSpawn					: LREAL;	// [s]
	lr_SpcSpawnInterval					: LREAL := 1;	// [s] random: the loop puts the products at an even pitch
	BeltPose							: ST_VisuPose;
	LatchPose							: ST_VisuPlanarPose;
	XtsPose								: ST_VisuPose;

	(* XTS loop: track position per mover *)
	b_SpcInitialised					: BOOL;
	lr_SpcS								: ARRAY[0..7] OF LREAL;	// [mm] per mover (n_SPC_MOVERS)
	n_SpcMode							: ARRAY[0..7] OF INT;
	udn_SpcProduct						: ARRAY[0..7] OF UDINT;	// [-] product pushed by the mover, 0 = none
	udn_SpcLastReleased					: UDINT;	// [-] product last handed back to the belt
	NoFingers							: ARRAY[0..VISU_GlobalConst_Param.VISU_un_MAX_FINGERS - 1] OF ST_VisuFingerState;
	un_Module							: UINT;	// [-] track module being set
	e_ModuleKind						: E_VisuModuleKind;
END_VAR
VAR CONSTANT
	(* Loop turned by 180 deg under the belt: its upper straight runs along MCS +X from X = 1000 to X = 4000, the
	   movers' tool points at the belt surface. *)
	lr_SPC_Y							: LREAL := 9000;	// [mm]
	lr_SPC_BELT_LENGTH					: LREAL := 5000;	// [mm]
	lr_SPC_BELT_SPEED					: LREAL := 150;	// [mm/s]
	(* Random gaps between arriving products. They stay above lr_SPC_SLOT, so a mover can always take the next
	   product over, and average lr_SPC_PITCH: the belt runs at the same speed on both sides, so the loop can only
	   even out the gaps, not change their mean. *)
	lr_SPC_MIN_GAP						: LREAL := 150;	// [mm]
	lr_SPC_GAP_SPREAD					: LREAL := 100;	// [mm] gaps lie between lr_SPC_MIN_GAP and lr_SPC_MIN_GAP + this
	lr_SPC_LOOP_END_X					: LREAL := 4000;	// [mm] MCS x of the loop origin, the downstream end
	un_SPC_STRAIGHT_MODULES				: UINT := 12;	// [-] straight XTS modules per side, joined at each end by two left curve modules
	lr_SPC_STRAIGHT						: LREAL := 3000;	// [mm] un_SPC_STRAIGHT_MODULES * 250
	lr_SPC_RADIUS						: LREAL := 159.15494309189535;	// [mm] two 250 mm quarter curves: 2 * 250 / pi
	lr_SPC_TOOL_OFFSET					: LREAL := 110;	// [mm] tool point outwards from the track: the belt surface
	n_SPC_MOVERS						: INT := 8;	// [-] size of the lr_SpcS, n_SpcMode and udn_SpcProduct arrays
	lr_SPC_SLOT							: LREAL := 130;	// [mm] queue spacing and minimum mover distance
	lr_SPC_TAKE_WINDOW					: LREAL := 40;	// [mm] take-over window from the start of the upper straight
	lr_SPC_PITCH						: LREAL := 200;	// [mm] constant product pitch on the outfeed
	lr_SPC_PUSH_SPEED					: LREAL := 450;	// [mm/s] maximum speed of a pushing mover
	lr_SPC_RETURN_SPEED					: LREAL := 900;	// [mm/s]
	lr_SPC_RELEASE_MIN_X				: LREAL := 2000;	// [mm] products are handed back to the belt from here...
	lr_SPC_RELEASE_MAX_X				: LREAL := 3800;	// [mm] ...up to here at the latest
	n_SPC_QUEUE							: INT := 0;
	n_SPC_PUSH							: INT := 1;
	n_SPC_RETURN						: INT := 2;
END_VAR

lr_Dt := DEMO_GlobalVar.DEMO_lr_Dt;


(****************************************************************************************************)
(* REGISTRATION (idempotent, every cycle)                                                           *)
(****************************************************************************************************)
fb_SpcBelt.m_Register(vio_Manifest := GVL_Visu.stManifest, vi_udn_Id := 13, vi_str_Name := 'Spacing belt');
fb_Spc.m_Register(vio_Manifest := GVL_Visu.stManifest, vi_udn_Id := 21, vi_str_Name := 'Spacer');


(****************************************************************************************************)
(* CONFIGURATION (idempotent, every cycle)                                                          *)
(****************************************************************************************************)
BeltPose.fX := 0;
BeltPose.fY := lr_SPC_Y;
BeltPose.fZ := DEMO_GlobalConst.DEMO_lr_BELT_Z;
fb_SpcBelt.m_SetPose(vi_Pose := BeltPose);
fb_SpcBelt.m_Configure(vi_lr_Length := lr_SPC_BELT_LENGTH, vi_lr_Width := DEMO_GlobalConst.DEMO_lr_BELT_WIDTH);
fb_SpcBelt.m_SetProductType(vi_udn_Id := 1, vi_lr_Length := DEMO_GlobalConst.DEMO_lr_PRODUCT_LENGTH,
	vi_lr_Width := DEMO_GlobalConst.DEMO_lr_PRODUCT_WIDTH, vi_lr_Height := DEMO_GlobalConst.DEMO_lr_PRODUCT_HEIGHT,
	vi_e_Shape := E_VisuProductShape.BOX, vi_lr_CornerRadius := 0);

(* Turned by 180 deg: the upper straight runs along MCS +X just below the belt, the tool points reach its surface. *)
XtsPose.fX := lr_SPC_LOOP_END_X;
XtsPose.fY := lr_SPC_Y;
XtsPose.fZ := DEMO_GlobalConst.DEMO_lr_BELT_Z - 2 * lr_SPC_RADIUS - lr_SPC_TOOL_OFFSET;
XtsPose.fRz := 180;
fb_Spc.m_SetPose(vi_Pose := XtsPose);
fb_Spc.m_Configure(vi_lr_ToolOffset := lr_SPC_TOOL_OFFSET, vi_lr_MoverLength := 100,
	vi_lr_MoverWidth := 60);
FOR un_Module := 1 TO 2 * (un_SPC_STRAIGHT_MODULES + 2) DO
	IF (un_Module - 1) MOD (un_SPC_STRAIGHT_MODULES + 2) < un_SPC_STRAIGHT_MODULES THEN
		e_ModuleKind := E_VisuModuleKind.STRAIGHT;
	ELSE
		e_ModuleKind := E_VisuModuleKind.CURVE_LEFT;
	END_IF
	fb_Spc.m_SetModule(vi_un_Module := un_Module, vi_e_Kind := e_ModuleKind,
		vi_lr_Length := VISU_GlobalConst.VISU_lr_XTS_MODULE_LENGTH);
END_FOR
fb_Spc.m_SetZone(vi_un_Zone := 1, vi_udn_ConveyorId := fb_SpcBelt.m_Id(),
	vi_lr_Start := lr_SPC_LOOP_END_X - lr_SPC_STRAIGHT, vi_lr_End := lr_SPC_LOOP_END_X - lr_SPC_STRAIGHT + lr_SPC_TAKE_WINDOW,
	vi_lr_AllocationOffset := 0, vi_lr_CcsOffset := lr_SPC_LOOP_END_X - lr_SPC_STRAIGHT,
	vi_lr_StartY := 0, vi_lr_EndY := 0);
fb_Spc.m_SetZone(vi_un_Zone := 2, vi_udn_ConveyorId := fb_SpcBelt.m_Id(),
	vi_lr_Start := lr_SPC_RELEASE_MIN_X, vi_lr_End := lr_SPC_RELEASE_MAX_X, vi_lr_AllocationOffset := 0,
	vi_lr_CcsOffset := lr_SPC_RELEASE_MIN_X, vi_lr_StartY := 0, vi_lr_EndY := 0);


(****************************************************************************************************)
(* BELT AND INFEED: random gaps                                                                     *)
(****************************************************************************************************)
lr_SpcBeltPosition := lr_SpcBeltPosition + lr_SPC_BELT_SPEED * lr_Dt;
fb_SpcBelt.m_SetBeltPosition(lr_SpcBeltPosition);
lr_SpcSinceSpawn := lr_SpcSinceSpawn + lr_Dt;
IF lr_SpcSinceSpawn >= lr_SpcSpawnInterval THEN
	lr_SpcSinceSpawn := 0;
	udn_Seed := udn_Seed * 1103515245 + 12345;
	lr_SpcSpawnInterval := (lr_SPC_MIN_GAP + UDINT_TO_LREAL(udn_Seed MOD 1000) / 1000.0 * lr_SPC_GAP_SPREAD)
							/ lr_SPC_BELT_SPEED;
	LatchPose.fX := 100;
	LatchPose.fY := lr_SPC_Y;
	LatchPose.fZ := DEMO_GlobalConst.DEMO_lr_BELT_Z;
	LatchPose.fRz := 0;
	IF fb_SpcBelt.m_LatchProduct(vi_udn_Id := DEMO_GlobalVar.DEMO_udn_NextId,
		vi_LatchPose := fb_SpcBelt.m_McsToBelt(vi_Pose := LatchPose),
		vi_udn_ProductType := 1, vi_lr_LatchBeltPosition := 0, vi_b_UseLatchBeltPosition := FALSE,
		vi_e_State := E_VisuProductState.DETECTED, vi_udn_ClientId := 0)
	THEN
		DEMO_GlobalVar.DEMO_udn_NextId := DEMO_GlobalVar.DEMO_udn_NextId + 1;
	END_IF
END_IF


(****************************************************************************************************)
(* XTS LOOP                                                                                         *)
(****************************************************************************************************)
m_Step();


(****************************************************************************************************)
(* HOUSEKEEPING                                                                                     *)
(****************************************************************************************************)
fb_SpcBelt.m_RemoveProductsBeyond(lr_SPC_BELT_LENGTH + DEMO_GlobalConst.DEMO_lr_REMOVE_BEYOND_END);

(****************************************************************************************************<br>
© Syntegon Group.<br>
All rights reserved, also regarding any disposal, exploitation, reproduction, editing, distribution,<br>
as well as in the event of applications for industrial property rights.<br>
*****************************************************************************************************<br>
DESCRIPTION:<br>
XTS loop under the belt: the queue head takes over the next product passing above the start of the upper<br>
straight and pushes it along the belt until it is lr_SPC_PITCH behind the product ahead, then lets the belt take<br>
it on and runs round to the queue.<br>
****************************************************************************************************)
METHOD PRIVATE m_Step : BOOL
VAR
	lr_TempPerimeter					: LREAL;	// [mm]
	lr_TempWait							: LREAL;	// [mm] track position of the start of the upper straight
	lr_TempStartX						: LREAL;	// [mm] MCS x of the start of the upper straight
	lr_TempX							: LREAL;	// [mm] MCS x
	lr_TempTarget						: LREAL;	// [mm] MCS x a pushing mover heads for
	lr_TempRef							: LREAL;	// [mm] MCS x of the product ahead
	lr_TempMinPush						: LREAL;	// [mm] track position of the last pushing mover
	n_TempI								: INT;
	n_TempJ								: INT;
	n_TempK								: INT;
	n_TempRank							: INT;
	n_TempHead							: INT;
	n_TempNext							: INT;
	n_TempIdx							: INT;
	un_TempIndex						: UINT;
	b_TempReady							: BOOL;
	b_TempDone							: ARRAY[0..7] OF BOOL;	// per mover (n_SPC_MOVERS)
	TempProduct							: ST_VisuProduct;
	TempPose							: ST_VisuPlanarPose;
	TempLatch							: ST_VisuPlanarPose;
END_VAR
(****************************************************************************************************)
(* QUEUE AND TAKE-OVER                                                                              *)
(****************************************************************************************************)
lr_TempPerimeter := fb_Spc.m_TrackLength();
lr_TempWait := lr_SPC_STRAIGHT + 3.141592653589793 * lr_SPC_RADIUS;
lr_TempStartX := lr_SPC_LOOP_END_X - lr_SPC_STRAIGHT;
IF NOT b_SpcInitialised THEN
	FOR n_TempI := 0 TO n_SPC_MOVERS - 1 DO
		lr_SpcS[n_TempI] := lr_TempWait - INT_TO_LREAL(n_TempI) * lr_SPC_SLOT;
		n_SpcMode[n_TempI] := n_SPC_QUEUE;
	END_FOR
	b_SpcInitialised := TRUE;
END_IF

(* Queued movers close up towards their slots before the start of the upper straight. *)
n_TempHead := -1;
FOR n_TempI := 0 TO n_SPC_MOVERS - 1 DO
	IF n_SpcMode[n_TempI] = n_SPC_QUEUE THEN
		n_TempRank := 0;
		FOR n_TempJ := 0 TO n_SPC_MOVERS - 1 DO
			IF n_SpcMode[n_TempJ] = n_SPC_QUEUE
			AND (lr_SpcS[n_TempJ] > lr_SpcS[n_TempI] OR (lr_SpcS[n_TempJ] = lr_SpcS[n_TempI] AND n_TempJ < n_TempI))
			THEN
				n_TempRank := n_TempRank + 1;
			END_IF
		END_FOR
		lr_SpcS[n_TempI] := MIN(lr_SpcS[n_TempI] + lr_SPC_RETURN_SPEED * lr_Dt,
								lr_TempWait - INT_TO_LREAL(n_TempRank) * lr_SPC_SLOT);
		IF n_TempRank = 0 THEN
			n_TempHead := n_TempI;
		END_IF
	END_IF
END_FOR

(* The ready queue head takes over the next product passing above the start of the upper straight, if the last
   pushing mover is at least one slot ahead. ST evaluates both operands of AND: test the head separately. *)
lr_TempMinPush := 1.0E9;
FOR n_TempI := 0 TO n_SPC_MOVERS - 1 DO
	IF n_SpcMode[n_TempI] = n_SPC_PUSH THEN
		lr_TempMinPush := MIN(lr_TempMinPush, lr_SpcS[n_TempI]);
	END_IF
END_FOR
b_TempReady := FALSE;
IF n_TempHead >= 0 THEN
	b_TempReady := lr_SpcS[n_TempHead] >= lr_TempWait - 1;
END_IF
IF b_TempReady THEN
	un_TempIndex := 0;
	WHILE n_SpcMode[n_TempHead] = n_SPC_QUEUE AND un_TempIndex < fb_SpcBelt.m_ProductCount() DO
		fb_SpcBelt.m_GetProduct(vi_un_Index := un_TempIndex, vo_Product => TempProduct, vo_Pose => TempPose);
		TempPose := fb_SpcBelt.m_BeltToMcs(vi_Pose := TempPose);
		lr_TempX := TempPose.fX - lr_TempStartX;
		IF TempProduct.eState = E_VisuProductState.DETECTED AND lr_TempX >= 0 AND lr_TempX < lr_SPC_TAKE_WINDOW
		AND lr_TempMinPush - lr_TempWait - lr_TempX >= lr_SPC_SLOT
		THEN
			fb_SpcBelt.m_SetProductState(vi_udn_Id := TempProduct.nId, vi_e_State := E_VisuProductState.ASSIGNED,
				vi_udn_ClientId := fb_Spc.m_Id(), vi_udn_MoverId := INT_TO_UDINT(n_TempHead + 1), vi_udn_FingerId := 0);
			udn_SpcProduct[n_TempHead] := TempProduct.nId;
			lr_SpcS[n_TempHead] := lr_TempWait + lr_TempX;
			n_SpcMode[n_TempHead] := n_SPC_PUSH;
		END_IF
		un_TempIndex := un_TempIndex + 1;
	END_WHILE
END_IF


(****************************************************************************************************)
(* PUSHING: the front mover first, so each one keeps the pitch to the product ahead of it            *)
(****************************************************************************************************)
lr_TempRef := 1.0E9;
IF udn_SpcLastReleased <> 0 THEN
	n_TempIdx := fb_SpcBelt.m_FindProduct(udn_SpcLastReleased);
	IF n_TempIdx >= 0 THEN
		fb_SpcBelt.m_GetProduct(vi_un_Index := INT_TO_UINT(n_TempIdx), vo_Product => TempProduct, vo_Pose => TempPose);
		TempPose := fb_SpcBelt.m_BeltToMcs(vi_Pose := TempPose);
		lr_TempRef := TempPose.fX;
	END_IF
END_IF
FOR n_TempI := 0 TO n_SPC_MOVERS - 1 DO
	b_TempDone[n_TempI] := n_SpcMode[n_TempI] <> n_SPC_PUSH;
END_FOR
FOR n_TempK := 1 TO n_SPC_MOVERS DO
	(* Next pushing mover: the one furthest along. *)
	n_TempNext := -1;
	FOR n_TempI := 0 TO n_SPC_MOVERS - 1 DO
		IF NOT b_TempDone[n_TempI] THEN
			IF n_TempNext < 0 THEN
				n_TempNext := n_TempI;
			ELSIF lr_SpcS[n_TempI] > lr_SpcS[n_TempNext] THEN
				n_TempNext := n_TempI;
			END_IF
		END_IF
	END_FOR
	IF n_TempNext < 0 THEN
		EXIT;
	END_IF
	b_TempDone[n_TempNext] := TRUE;

	n_TempIdx := fb_SpcBelt.m_FindProduct(udn_SpcProduct[n_TempNext]);
	IF n_TempIdx < 0 THEN
		(* The product is gone: run round to the queue. *)
		udn_SpcProduct[n_TempNext] := 0;
		n_SpcMode[n_TempNext] := n_SPC_RETURN;
	ELSE
		lr_TempX := lr_TempStartX + lr_SpcS[n_TempNext] - lr_TempWait;
		lr_TempTarget := MIN(lr_SPC_RELEASE_MAX_X, lr_TempRef - lr_SPC_PITCH);
		lr_TempX := lr_TempX + LIMIT(0, lr_TempTarget - lr_TempX, lr_SPC_PUSH_SPEED * lr_Dt);
		lr_SpcS[n_TempNext] := lr_TempWait + lr_TempX - lr_TempStartX;
		TempLatch.fX := lr_TempX;
		TempLatch.fY := lr_SPC_Y;
		TempLatch.fZ := DEMO_GlobalConst.DEMO_lr_BELT_Z;
		TempLatch.fRz := 0;
		fb_SpcBelt.m_MoveProduct(vi_udn_Id := udn_SpcProduct[n_TempNext],
			vi_Pose := fb_SpcBelt.m_McsToBelt(vi_Pose := TempLatch));
		lr_TempRef := lr_TempX;

		(* At the pitch behind the product ahead (or at the end of the release area): the belt takes it on. Only the
		   front mover lets go, so a returning mover never overtakes one that still pushes. *)
		IF n_TempK = 1 AND lr_TempX >= lr_SPC_RELEASE_MIN_X AND ABS(lr_TempTarget - lr_TempX) < 0.5 THEN
			(* Put back onto the belt by the loop: PLACED, so it does not count as missed at the belt end. *)
			fb_SpcBelt.m_SetProductState(vi_udn_Id := udn_SpcProduct[n_TempNext], vi_e_State := E_VisuProductState.PLACED,
				vi_udn_ClientId := fb_Spc.m_Id(), vi_udn_MoverId := 0, vi_udn_FingerId := 0);
			udn_SpcLastReleased := udn_SpcProduct[n_TempNext];
			udn_SpcProduct[n_TempNext] := 0;
			n_SpcMode[n_TempNext] := n_SPC_RETURN;
		END_IF
	END_IF
END_FOR


(****************************************************************************************************)
(* RETURN AND REPORT                                                                                *)
(****************************************************************************************************)
fb_Spc.m_SetMoverCount(INT_TO_UINT(n_SPC_MOVERS));
FOR n_TempI := 0 TO n_SPC_MOVERS - 1 DO
	(* Back along the lower straight; past the perimeter the mover joins the queue. *)
	IF n_SpcMode[n_TempI] = n_SPC_RETURN THEN
		lr_SpcS[n_TempI] := lr_SpcS[n_TempI] + lr_SPC_RETURN_SPEED * lr_Dt;
		IF lr_SpcS[n_TempI] >= lr_TempPerimeter THEN
			lr_SpcS[n_TempI] := lr_SpcS[n_TempI] - lr_TempPerimeter;
			n_SpcMode[n_TempI] := n_SPC_QUEUE;
		END_IF
	END_IF
	fb_Spc.m_SetMover(vi_un_Index := INT_TO_UINT(n_TempI), vi_udn_Id := INT_TO_UDINT(n_TempI + 1),
		vi_lr_Position := lr_SpcS[n_TempI], vi_FingerStates := NoFingers, vi_b_Fault := FALSE, vi_str_FaultMessage := '');
END_FOR
m_Step := TRUE;
END_METHOD

END_PROGRAM

// ---- POUs/P_VisuDemoStress.TcPOU
(****************************************************************************************************<br>
© Syntegon Group.<br>
All rights reserved, also regarding any disposal, exploitation, reproduction, editing, distribution,<br>
as well as in the event of applications for industrial property rights.<br>
*****************************************************************************************************<br>
DESCRIPTION:<br>
DEMO ONLY: load test (Y = 11000), off unless DEMO_GlobalVar.DEMO_un_StressProducts is set online. A wide stress<br>
belt carries that many products in lanes (at most VISU_un_MAX_PRODUCTS less four rows): it fills up within a few<br>
seconds, then a row enters at its start every pitch and leaves beyond its end, and one product per row is<br>
rejected halfway (m_SetProductState on a full register). It measures the task's execution time, so the cost of<br>
large registers in the library shows in udn_MaxExecTime, and the gateway's /health shows whether the gateway reads<br>
registers the PLC is rearranging (duplicateProducts, flickeringProducts). Called by P_VisuDemo.<br>
****************************************************************************************************)
PROGRAM P_VisuDemoStress
VAR
	fb_StressBelt						: _FB_VisuConveyor;
	b_Registered						: BOOL;	// the stress belt is in the manifest
	b_On								: BOOL;	// DEMO_un_StressProducts was above 0 in the previous cycle

	(* Belt *)
	lr_Dt								: LREAL;	// [s] cycle time
	un_Target							: UINT;	// [-] products asked for, limited to the register
	un_Rows								: UINT;	// [-] rows of products along the belt
	lr_BeltLength						: LREAL;	// [mm]
	lr_BeltPosition						: LREAL;	// [mm]
	lr_EntryStart						: LREAL;	// [mm] belt position when the first row entered
	lr_NextRow							: LREAL;	// [mm] belt position at which the next row enters
	udn_RowCount						: UDINT;	// [-] rows entered at the start so far
	udn_RowFirstId						: ARRAY[0..VISU_GlobalConst_Param.VISU_un_MAX_PRODUCTS / 10] OF UDINT;	// [-] id of the first product per entered row, a ring (un_STRESS_LANES lanes)
	un_FillRow							: UINT;	// [-] rows filled in from the belt end since the length changed
	un_FilledNow						: UINT;	// [-] rows filled in this cycle
	BeltPose							: ST_VisuPose;

	(* Measurements, read them online *)
	dn_TaskIndex						: DINT;
	udn_LastExecTime					: UDINT;	// [100 ns] last cycle of the calling task, all programs
	udn_MaxExecTime						: UDINT;	// [100 ns] largest udn_LastExecTime since the last reset
	udn_ExceededCount					: UDINT;	// [-] cycles that exceeded the task cycle time since the last reset
	b_ResetMax							: BOOL;	// TRUE: restart udn_MaxExecTime and udn_ExceededCount
	un_Products							: UINT;	// [-] products in the stress belt's register
END_VAR
VAR CONSTANT
	lr_STRESS_Y							: LREAL := 11000;	// [mm]
	un_STRESS_LANES						: UINT := 10;	// [-] also the divisor of the udn_RowFirstId size
	lr_STRESS_LANE_WIDTH				: LREAL := 100;	// [mm]
	lr_STRESS_PITCH						: LREAL := 150;	// [mm] distance between two rows along the belt
	lr_STRESS_SPEED						: LREAL := 300;	// [mm/s]
	un_STRESS_FILL_ROWS					: UINT := 2;	// [-] rows filled in per cycle while the belt fills up
END_VAR

lr_Dt := DEMO_GlobalVar.DEMO_lr_Dt;


(****************************************************************************************************)
(* TASK LOAD                                                                                        *)
(****************************************************************************************************)
dn_TaskIndex := Tc2_System.GETCURTASKINDEXEX();
IF dn_TaskIndex > 0 THEN
	IF b_ResetMax THEN
		b_ResetMax := FALSE;
		udn_MaxExecTime := 0;
		udn_ExceededCount := 0;
	END_IF
	udn_LastExecTime := TwinCAT_SystemInfoVarList._TaskInfo[dn_TaskIndex].LastExecTime;
	udn_MaxExecTime := MAX(udn_MaxExecTime, udn_LastExecTime);
	IF TwinCAT_SystemInfoVarList._TaskInfo[dn_TaskIndex].CycleTimeExceeded THEN
		udn_ExceededCount := udn_ExceededCount + 1;
	END_IF
END_IF


(****************************************************************************************************)
(* REGISTRATION AND CONFIGURATION: only once a load is asked for                                    *)
(****************************************************************************************************)
un_Target := MIN(DEMO_GlobalVar.DEMO_un_StressProducts, VISU_GlobalConst_Param.VISU_un_MAX_PRODUCTS - 4 * un_STRESS_LANES);
IF un_Target = 0 AND NOT b_Registered THEN
	RETURN;
END_IF
fb_StressBelt.m_Register(vio_Manifest := GVL_Visu.stManifest, vi_udn_Id := 14, vi_str_Name := 'Stress belt');
IF NOT b_Registered THEN
	b_Registered := TRUE;
	lr_EntryStart := lr_BeltPosition;
	lr_NextRow := lr_BeltPosition;
END_IF

(* Set back to 0 the belt keeps its length and runs empty. *)
IF un_Target > 0 AND (un_Target + un_STRESS_LANES - 1) / un_STRESS_LANES <> un_Rows THEN
	un_Rows := (un_Target + un_STRESS_LANES - 1) / un_STRESS_LANES;
	(* The entering rows have covered at most the old length: a longer belt is filled in beyond it. *)
	lr_EntryStart := lr_BeltPosition - MIN(lr_BeltLength, lr_BeltPosition - lr_EntryStart);
	lr_BeltLength := UINT_TO_LREAL(un_Rows) * lr_STRESS_PITCH;
	un_FillRow := 0;
END_IF
BeltPose.fX := 0;
BeltPose.fY := lr_STRESS_Y;
BeltPose.fZ := DEMO_GlobalConst.DEMO_lr_BELT_Z;
fb_StressBelt.m_SetPose(vi_Pose := BeltPose);
fb_StressBelt.m_Configure(vi_lr_Length := lr_BeltLength,
	vi_lr_Width := UINT_TO_LREAL(un_STRESS_LANES) * lr_STRESS_LANE_WIDTH + 100);
fb_StressBelt.m_SetProductType(vi_udn_Id := 1, vi_lr_Length := DEMO_GlobalConst.DEMO_lr_PRODUCT_LENGTH,
	vi_lr_Width := DEMO_GlobalConst.DEMO_lr_PRODUCT_WIDTH, vi_lr_Height := DEMO_GlobalConst.DEMO_lr_PRODUCT_HEIGHT,
	vi_e_Shape := E_VisuProductShape.BOX, vi_lr_CornerRadius := 0);


(****************************************************************************************************)
(* BELT: fill up from the end, then a row enters at the start every pitch                           *)
(****************************************************************************************************)
lr_BeltPosition := lr_BeltPosition + lr_STRESS_SPEED * lr_Dt;
fb_StressBelt.m_SetBeltPosition(lr_BeltPosition);

(* Switched on: start from an empty belt and fill it up, so a measurement always gets the load asked for. *)
IF DEMO_GlobalVar.DEMO_un_StressProducts > 0 AND NOT b_On THEN
	fb_StressBelt.m_RemoveProductsBeyond(-1.0E12);
	lr_EntryStart := lr_BeltPosition;
	lr_NextRow := lr_BeltPosition;
	un_FillRow := 0;
END_IF
b_On := DEMO_GlobalVar.DEMO_un_StressProducts > 0;

